    PROC Decorar_Ing165(PERS wobjdata WO_Pastel)
        Mover_en_vacio;
        MoveJ Target_Home_10,Vel_Vacio_Rap,Z_Vacio_Rap,Prototipo_JSDaleman\WObj:=wobj0;
        ReiniciarIndices;
        path_contacto_actual:="p_contacto_165";
        path_vacio_actual:="p_vacio_165";
        Path_Tapa_165ing WO_Pastel;
        Mover_en_vacio;
        MoveJ Target_Home_10,Vel_Vacio_Rap,Z_Vacio_Rap,Prototipo_JSDaleman\WObj:=wobj0;
    ENDPROC
    PROC Path_Tapa_165ing(PERS wobjdata WO_Pastel)
        Path_vacio_ejecucion p_vacio_165, 1, WO_Pastel, FALSE;
        Path_contacto_ejecucion p_contacto_165, 1, 7, WO_Pastel, TRUE;
        Path_vacio_ejecucion p_vacio_165, 2, WO_Pastel, FALSE;
        index_vacio_destino:=15;
        Path_contacto_ejecucion p_contacto_165, 8, 10, WO_Pastel, FALSE;
        Mover_en_contacto;
        TriggC p_contacto_165{11},p_contacto_165{12},Vel_Proceso,triggContactoCir,Z_Proceso,Prototipo_JSDaleman\WObj:=WO_Pastel;
        TriggC p_contacto_165{13},p_contacto_165{14},Vel_Proceso,triggContactoCir,Z_Proceso,Prototipo_JSDaleman\WObj:=WO_Pastel;
        Mover_a_vacio;
        TriggL p_contacto_165{15},Vel_Acercamiento,triggContacto,Z_Acercamiento,Prototipo_JSDaleman\WObj:=WO_Pastel;
        Path_vacio_ejecucion p_vacio_165, 3, WO_Pastel, FALSE;
        index_vacio_destino:=21;
        Mover_a_contacto;
        TriggL p_contacto_165{16},Vel_Acercamiento,triggContacto,Z_Acercamiento,Prototipo_JSDaleman\WObj:=WO_Pastel;
        Mover_en_contacto;
        TriggC p_contacto_165{17},p_contacto_165{18},Vel_Proceso,triggContactoCir,Z_Proceso,Prototipo_JSDaleman\WObj:=WO_Pastel;
        TriggC p_contacto_165{19},p_contacto_165{20},Vel_Proceso,triggContactoCir,Z_Proceso,Prototipo_JSDaleman\WObj:=WO_Pastel;
        Mover_a_vacio;
        TriggL p_contacto_165{21},Vel_Acercamiento,triggContacto,Z_Acercamiento,Prototipo_JSDaleman\WObj:=WO_Pastel;
        Path_vacio_ejecucion p_vacio_165, 4, WO_Pastel, FALSE;
        index_vacio_destino:=28;
        Path_contacto_ejecucion p_contacto_165, 22, 23, WO_Pastel, FALSE;
        Mover_en_contacto;
        TriggC p_contacto_165{24},p_contacto_165{25},Vel_Proceso,triggContactoCir,Z_Proceso,Prototipo_JSDaleman\WObj:=WO_Pastel;
        TriggL p_contacto_165{26},Vel_Proceso,triggContacto,Z_Proceso,Prototipo_JSDaleman\WObj:=WO_Pastel;
        TriggL p_contacto_165{27},Vel_Proceso,triggContacto,Z_Proceso,Prototipo_JSDaleman\WObj:=WO_Pastel;
        Mover_a_vacio;
        TriggL p_contacto_165{28},Vel_Acercamiento,triggContacto,Z_Acercamiento,Prototipo_JSDaleman\WObj:=WO_Pastel;
        Path_vacio_ejecucion p_vacio_165, 5, WO_Pastel, FALSE;
        Path_contacto_ejecucion p_contacto_165, 29, 31, WO_Pastel, TRUE;
        Path_vacio_ejecucion p_vacio_165, 6, WO_Pastel, FALSE;
        Path_contacto_ejecucion p_contacto_165, 32, 39, WO_Pastel, TRUE;
        Path_vacio_ejecucion p_vacio_165, 7, WO_Pastel, FALSE;
        index_vacio_destino:=47;
        Path_contacto_ejecucion p_contacto_165, 40, 42, WO_Pastel, FALSE;
        Mover_en_contacto;
        TriggC p_contacto_165{43},p_contacto_165{44},Vel_Proceso,triggContactoCir,Z_Proceso,Prototipo_JSDaleman\WObj:=WO_Pastel;
        TriggC p_contacto_165{45},p_contacto_165{46},Vel_Proceso,triggContactoCir,Z_Proceso,Prototipo_JSDaleman\WObj:=WO_Pastel;
        Mover_a_vacio;
        TriggL p_contacto_165{47},Vel_Acercamiento,triggContacto,Z_Acercamiento,Prototipo_JSDaleman\WObj:=WO_Pastel;
        Path_vacio_ejecucion p_vacio_165, 8, WO_Pastel, FALSE;
        index_vacio_destino:=55;
        Path_contacto_ejecucion p_contacto_165, 48, 50, WO_Pastel, FALSE;
        Mover_en_contacto;
        TriggC p_contacto_165{51},p_contacto_165{52},Vel_Proceso,triggContactoCir,Z_Proceso,Prototipo_JSDaleman\WObj:=WO_Pastel;
        TriggC p_contacto_165{53},p_contacto_165{54},Vel_Proceso,triggContactoCir,Z_Proceso,Prototipo_JSDaleman\WObj:=WO_Pastel;
        Mover_a_vacio;
        TriggL p_contacto_165{55},Vel_Acercamiento,triggContacto,Z_Acercamiento,Prototipo_JSDaleman\WObj:=WO_Pastel;
        Path_vacio_ejecucion p_vacio_165, 9, WO_Pastel, FALSE;
        index_vacio_destino:=63;
        Path_contacto_ejecucion p_contacto_165, 56, 58, WO_Pastel, FALSE;
        Mover_en_contacto;
        TriggC p_contacto_165{59},p_contacto_165{60},Vel_Proceso,triggContactoCir,Z_Proceso,Prototipo_JSDaleman\WObj:=WO_Pastel;
        TriggC p_contacto_165{61},p_contacto_165{62},Vel_Proceso,triggContactoCir,Z_Proceso,Prototipo_JSDaleman\WObj:=WO_Pastel;
        Mover_a_vacio;
        TriggL p_contacto_165{63},Vel_Acercamiento,triggContacto,Z_Acercamiento,Prototipo_JSDaleman\WObj:=WO_Pastel;
        Path_vacio_ejecucion p_vacio_165, 10, WO_Pastel, FALSE;
        index_vacio_destino:=70;
        Mover_a_contacto;
        TriggL p_contacto_165{64},Vel_Acercamiento,triggContacto,Z_Acercamiento,Prototipo_JSDaleman\WObj:=WO_Pastel;
        Mover_en_contacto;
        TriggC p_contacto_165{65},p_contacto_165{66},Vel_Proceso,triggContactoCir,Z_Proceso,Prototipo_JSDaleman\WObj:=WO_Pastel;
        TriggC p_contacto_165{67},p_contacto_165{68},Vel_Proceso,triggContactoCir,Z_Proceso,Prototipo_JSDaleman\WObj:=WO_Pastel;
        TriggL p_contacto_165{69},Vel_Proceso,triggContacto,Z_Proceso,Prototipo_JSDaleman\WObj:=WO_Pastel;
        Mover_a_vacio;
        TriggL p_contacto_165{70},Vel_Acercamiento,triggContacto,Z_Acercamiento,Prototipo_JSDaleman\WObj:=WO_Pastel;
        Path_vacio_ejecucion p_vacio_165, 11, WO_Pastel, FALSE;
        Path_contacto_ejecucion p_contacto_165, 71, 73, WO_Pastel, TRUE;
        Path_vacio_ejecucion p_vacio_165, 12, WO_Pastel, FALSE;
        index_vacio_destino:=80;
        Path_contacto_ejecucion p_contacto_165, 74, 76, WO_Pastel, FALSE;
        Mover_en_contacto;
        TriggC p_contacto_165{77},p_contacto_165{78},Vel_Proceso,triggContactoCir,Z_Proceso,Prototipo_JSDaleman\WObj:=WO_Pastel;
        TriggL p_contacto_165{79},Vel_Proceso,triggContacto,Z_Proceso,Prototipo_JSDaleman\WObj:=WO_Pastel;
        Mover_a_vacio;
        TriggL p_contacto_165{80},Vel_Acercamiento,triggContacto,Z_Acercamiento,Prototipo_JSDaleman\WObj:=WO_Pastel;
        Path_vacio_ejecucion p_vacio_165, 13, WO_Pastel, FALSE;
        index_vacio_destino:=90;
        Mover_a_contacto;
        TriggL p_contacto_165{81},Vel_Acercamiento,triggContacto,Z_Acercamiento,Prototipo_JSDaleman\WObj:=WO_Pastel;
        Mover_en_contacto;
        TriggC p_contacto_165{82},p_contacto_165{83},Vel_Proceso,triggContactoCir,Z_Proceso,Prototipo_JSDaleman\WObj:=WO_Pastel;
        TriggL p_contacto_165{84},Vel_Proceso,triggContacto,Z_Proceso,Prototipo_JSDaleman\WObj:=WO_Pastel;
        TriggL p_contacto_165{85},Vel_Proceso,triggContacto,Z_Proceso,Prototipo_JSDaleman\WObj:=WO_Pastel;
        TriggC p_contacto_165{86},p_contacto_165{87},Vel_Proceso,triggContactoCir,Z_Proceso,Prototipo_JSDaleman\WObj:=WO_Pastel;
        TriggC p_contacto_165{88},p_contacto_165{89},Vel_Proceso,triggContactoCir,Z_Proceso,Prototipo_JSDaleman\WObj:=WO_Pastel;
        Mover_a_vacio;
        TriggL p_contacto_165{90},Vel_Acercamiento,triggContacto,Z_Acercamiento,Prototipo_JSDaleman\WObj:=WO_Pastel;
        Path_vacio_ejecucion p_vacio_165, 14, WO_Pastel, FALSE;
        index_vacio_destino:=97;
        Mover_a_contacto;
        TriggL p_contacto_165{91},Vel_Acercamiento,triggContacto,Z_Acercamiento,Prototipo_JSDaleman\WObj:=WO_Pastel;
        Mover_en_contacto;
        TriggC p_contacto_165{92},p_contacto_165{93},Vel_Proceso,triggContactoCir,Z_Proceso,Prototipo_JSDaleman\WObj:=WO_Pastel;
        TriggC p_contacto_165{94},p_contacto_165{95},Vel_Proceso,triggContactoCir,Z_Proceso,Prototipo_JSDaleman\WObj:=WO_Pastel;
        TriggL p_contacto_165{96},Vel_Proceso,triggContacto,Z_Proceso,Prototipo_JSDaleman\WObj:=WO_Pastel;
        Mover_a_vacio;
        TriggL p_contacto_165{97},Vel_Acercamiento,triggContacto,Z_Acercamiento,Prototipo_JSDaleman\WObj:=WO_Pastel;
        Path_vacio_ejecucion p_vacio_165, 15, WO_Pastel, FALSE;
        index_vacio_destino:=104;
        Path_contacto_ejecucion p_contacto_165, 98, 100, WO_Pastel, FALSE;
        Mover_en_contacto;
        TriggC p_contacto_165{101},p_contacto_165{102},Vel_Proceso,triggContactoCir,Z_Proceso,Prototipo_JSDaleman\WObj:=WO_Pastel;
        TriggL p_contacto_165{103},Vel_Proceso,triggContacto,Z_Proceso,Prototipo_JSDaleman\WObj:=WO_Pastel;
        Mover_a_vacio;
        TriggL p_contacto_165{104},Vel_Acercamiento,triggContacto,Z_Acercamiento,Prototipo_JSDaleman\WObj:=WO_Pastel;
        Path_vacio_ejecucion p_vacio_165, 16, WO_Pastel, FALSE;
        Path_contacto_ejecucion p_contacto_165, 105, 107, WO_Pastel, TRUE;
        Path_vacio_ejecucion p_vacio_165, 17, WO_Pastel, FALSE;
        Path_contacto_ejecucion p_contacto_165, 108, 109, WO_Pastel, TRUE;
        Path_vacio_ejecucion p_vacio_165, 18, WO_Pastel, FALSE;
        index_vacio_destino:=116;
        Mover_a_contacto;
        TriggL p_contacto_165{110},Vel_Acercamiento,triggContacto,Z_Acercamiento,Prototipo_JSDaleman\WObj:=WO_Pastel;
        Mover_en_contacto;
        TriggC p_contacto_165{111},p_contacto_165{112},Vel_Proceso,triggContactoCir,Z_Proceso,Prototipo_JSDaleman\WObj:=WO_Pastel;
        TriggC p_contacto_165{113},p_contacto_165{114},Vel_Proceso,triggContactoCir,Z_Proceso,Prototipo_JSDaleman\WObj:=WO_Pastel;
        TriggL p_contacto_165{115},Vel_Proceso,triggContacto,Z_Proceso,Prototipo_JSDaleman\WObj:=WO_Pastel;
        Mover_a_vacio;
        TriggL p_contacto_165{116},Vel_Acercamiento,triggContacto,Z_Acercamiento,Prototipo_JSDaleman\WObj:=WO_Pastel;
        Path_vacio_ejecucion p_vacio_165, 19, WO_Pastel, FALSE;
        Path_contacto_ejecucion p_contacto_165, 117, 121, WO_Pastel, TRUE;
        Path_vacio_ejecucion p_vacio_165, 20, WO_Pastel, FALSE;
        Path_contacto_ejecucion p_contacto_165, 122, 124, WO_Pastel, TRUE;
        Path_vacio_ejecucion p_vacio_165, 21, WO_Pastel, FALSE;
        Path_contacto_ejecucion p_contacto_165, 125, 127, WO_Pastel, TRUE;
        Path_vacio_ejecucion p_vacio_165, 22, WO_Pastel, FALSE;
        index_vacio_destino:=135;
        Path_contacto_ejecucion p_contacto_165, 128, 130, WO_Pastel, FALSE;
        Mover_en_contacto;
        TriggC p_contacto_165{131},p_contacto_165{132},Vel_Proceso,triggContactoCir,Z_Proceso,Prototipo_JSDaleman\WObj:=WO_Pastel;
        TriggC p_contacto_165{133},p_contacto_165{134},Vel_Proceso,triggContactoCir,Z_Proceso,Prototipo_JSDaleman\WObj:=WO_Pastel;
        Mover_a_vacio;
        TriggL p_contacto_165{135},Vel_Acercamiento,triggContacto,Z_Acercamiento,Prototipo_JSDaleman\WObj:=WO_Pastel;
        Path_vacio_ejecucion p_vacio_165, 23, WO_Pastel, FALSE;
        index_vacio_destino:=139;
        Mover_a_contacto;
        TriggL p_contacto_165{136},Vel_Acercamiento,triggContacto,Z_Acercamiento,Prototipo_JSDaleman\WObj:=WO_Pastel;
        Mover_en_contacto;
        TriggC p_contacto_165{137},p_contacto_165{138},Vel_Proceso,triggContactoCir,Z_Proceso,Prototipo_JSDaleman\WObj:=WO_Pastel;
        Mover_a_vacio;
        TriggL p_contacto_165{139},Vel_Acercamiento,triggContacto,Z_Acercamiento,Prototipo_JSDaleman\WObj:=WO_Pastel;
        Path_vacio_ejecucion p_vacio_165, 24, WO_Pastel, FALSE;
        index_vacio_destino:=143;
        Mover_a_contacto;
        TriggL p_contacto_165{140},Vel_Acercamiento,triggContacto,Z_Acercamiento,Prototipo_JSDaleman\WObj:=WO_Pastel;
        Mover_en_contacto;
        TriggC p_contacto_165{141},p_contacto_165{142},Vel_Proceso,triggContactoCir,Z_Proceso,Prototipo_JSDaleman\WObj:=WO_Pastel;
        Mover_a_vacio;
        TriggL p_contacto_165{143},Vel_Acercamiento,triggContacto,Z_Acercamiento,Prototipo_JSDaleman\WObj:=WO_Pastel;
        Path_vacio_ejecucion p_vacio_165, 25, WO_Pastel, FALSE;
        index_vacio_destino:=147;
        Mover_a_contacto;
        TriggL p_contacto_165{144},Vel_Acercamiento,triggContacto,Z_Acercamiento,Prototipo_JSDaleman\WObj:=WO_Pastel;
        Mover_en_contacto;
        TriggC p_contacto_165{145},p_contacto_165{146},Vel_Proceso,triggContactoCir,Z_Proceso,Prototipo_JSDaleman\WObj:=WO_Pastel;
        Mover_a_vacio;
        TriggL p_contacto_165{147},Vel_Acercamiento,triggContacto,Z_Acercamiento,Prototipo_JSDaleman\WObj:=WO_Pastel;
        Path_vacio_ejecucion p_vacio_165, 26, WO_Pastel, FALSE;
        Path_contacto_ejecucion p_contacto_165, 148, 150, WO_Pastel, TRUE;
        Path_vacio_ejecucion p_vacio_165, 27, WO_Pastel, FALSE;
        index_vacio_destino:=154;
        Mover_a_contacto;
        TriggL p_contacto_165{151},Vel_Acercamiento,triggContacto,Z_Acercamiento,Prototipo_JSDaleman\WObj:=WO_Pastel;
        Mover_en_contacto;
        TriggC p_contacto_165{152},p_contacto_165{153},Vel_Proceso,triggContactoCir,Z_Proceso,Prototipo_JSDaleman\WObj:=WO_Pastel;
        Mover_a_vacio;
        TriggL p_contacto_165{154},Vel_Acercamiento,triggContacto,Z_Acercamiento,Prototipo_JSDaleman\WObj:=WO_Pastel;
        Path_vacio_ejecucion p_vacio_165, 28, WO_Pastel, FALSE;
        index_vacio_destino:=158;
        Mover_a_contacto;
        TriggL p_contacto_165{155},Vel_Acercamiento,triggContacto,Z_Acercamiento,Prototipo_JSDaleman\WObj:=WO_Pastel;
        Mover_en_contacto;
        TriggC p_contacto_165{156},p_contacto_165{157},Vel_Proceso,triggContactoCir,Z_Proceso,Prototipo_JSDaleman\WObj:=WO_Pastel;
        Mover_a_vacio;
        TriggL p_contacto_165{158},Vel_Acercamiento,triggContacto,Z_Acercamiento,Prototipo_JSDaleman\WObj:=WO_Pastel;
        Path_vacio_ejecucion p_vacio_165, 29, WO_Pastel, FALSE;
        index_vacio_destino:=162;
        Mover_a_contacto;
        TriggL p_contacto_165{159},Vel_Acercamiento,triggContacto,Z_Acercamiento,Prototipo_JSDaleman\WObj:=WO_Pastel;
        Mover_en_contacto;
        TriggC p_contacto_165{160},p_contacto_165{161},Vel_Proceso,triggContactoCir,Z_Proceso,Prototipo_JSDaleman\WObj:=WO_Pastel;
        Mover_a_vacio;
        TriggL p_contacto_165{162},Vel_Acercamiento,triggContacto,Z_Acercamiento,Prototipo_JSDaleman\WObj:=WO_Pastel;
        Path_vacio_ejecucion p_vacio_165, 30, WO_Pastel, FALSE;
        index_vacio_destino:=170;
        Path_contacto_ejecucion p_contacto_165, 163, 165, WO_Pastel, FALSE;
        Mover_en_contacto;
        TriggC p_contacto_165{166},p_contacto_165{167},Vel_Proceso,triggContactoCir,Z_Proceso,Prototipo_JSDaleman\WObj:=WO_Pastel;
        TriggC p_contacto_165{168},p_contacto_165{169},Vel_Proceso,triggContactoCir,Z_Proceso,Prototipo_JSDaleman\WObj:=WO_Pastel;
        Mover_a_vacio;
        TriggL p_contacto_165{170},Vel_Acercamiento,triggContacto,Z_Acercamiento,Prototipo_JSDaleman\WObj:=WO_Pastel;
        Path_vacio_ejecucion p_vacio_165, 31, WO_Pastel, FALSE;
        index_vacio_destino:=178;
        Path_contacto_ejecucion p_contacto_165, 171, 173, WO_Pastel, FALSE;
        Mover_en_contacto;
        TriggC p_contacto_165{174},p_contacto_165{175},Vel_Proceso,triggContactoCir,Z_Proceso,Prototipo_JSDaleman\WObj:=WO_Pastel;
        TriggL p_contacto_165{176},Vel_Proceso,triggContacto,Z_Proceso,Prototipo_JSDaleman\WObj:=WO_Pastel;
        TriggL p_contacto_165{177},Vel_Proceso,triggContacto,Z_Proceso,Prototipo_JSDaleman\WObj:=WO_Pastel;
        Mover_a_vacio;
        TriggL p_contacto_165{178},Vel_Acercamiento,triggContacto,Z_Acercamiento,Prototipo_JSDaleman\WObj:=WO_Pastel;
        Path_vacio_ejecucion p_vacio_165, 32, WO_Pastel, FALSE;
        index_vacio_destino:=184;
        Mover_a_contacto;
        TriggL p_contacto_165{179},Vel_Acercamiento,triggContacto,Z_Acercamiento,Prototipo_JSDaleman\WObj:=WO_Pastel;
        Mover_en_contacto;
        TriggC p_contacto_165{180},p_contacto_165{181},Vel_Proceso,triggContactoCir,Z_Proceso,Prototipo_JSDaleman\WObj:=WO_Pastel;
        TriggC p_contacto_165{182},p_contacto_165{183},Vel_Proceso,triggContactoCir,Z_Proceso,Prototipo_JSDaleman\WObj:=WO_Pastel;
        Mover_a_vacio;
        TriggL p_contacto_165{184},Vel_Acercamiento,triggContacto,Z_Acercamiento,Prototipo_JSDaleman\WObj:=WO_Pastel;
        Path_vacio_ejecucion p_vacio_165, 33, WO_Pastel, FALSE;
        index_vacio_destino:=190;
        Mover_a_contacto;
        TriggL p_contacto_165{185},Vel_Acercamiento,triggContacto,Z_Acercamiento,Prototipo_JSDaleman\WObj:=WO_Pastel;
        Mover_en_contacto;
        TriggC p_contacto_165{186},p_contacto_165{187},Vel_Proceso,triggContactoCir,Z_Proceso,Prototipo_JSDaleman\WObj:=WO_Pastel;
        TriggC p_contacto_165{188},p_contacto_165{189},Vel_Proceso,triggContactoCir,Z_Proceso,Prototipo_JSDaleman\WObj:=WO_Pastel;
        Mover_a_vacio;
        TriggL p_contacto_165{190},Vel_Acercamiento,triggContacto,Z_Acercamiento,Prototipo_JSDaleman\WObj:=WO_Pastel;
        Path_vacio_ejecucion p_vacio_165, 34, WO_Pastel, FALSE;
        index_vacio_destino:=198;
        Mover_a_contacto;
        TriggL p_contacto_165{191},Vel_Acercamiento,triggContacto,Z_Acercamiento,Prototipo_JSDaleman\WObj:=WO_Pastel;
        Mover_en_contacto;
        TriggC p_contacto_165{192},p_contacto_165{193},Vel_Proceso,triggContactoCir,Z_Proceso,Prototipo_JSDaleman\WObj:=WO_Pastel;
        TriggL p_contacto_165{194},Vel_Proceso,triggContacto,Z_Proceso,Prototipo_JSDaleman\WObj:=WO_Pastel;
        TriggL p_contacto_165{195},Vel_Proceso,triggContacto,Z_Proceso,Prototipo_JSDaleman\WObj:=WO_Pastel;
        TriggC p_contacto_165{196},p_contacto_165{197},Vel_Proceso,triggContactoCir,Z_Proceso,Prototipo_JSDaleman\WObj:=WO_Pastel;
        Mover_a_vacio;
        TriggL p_contacto_165{198},Vel_Acercamiento,triggContacto,Z_Acercamiento,Prototipo_JSDaleman\WObj:=WO_Pastel;
        Path_vacio_ejecucion p_vacio_165, 35, WO_Pastel, FALSE;
        Path_contacto_ejecucion p_contacto_165, 199, 201, WO_Pastel, TRUE;
        Path_vacio_ejecucion p_vacio_165, 36, WO_Pastel, FALSE;
        Path_contacto_ejecucion p_contacto_165, 202, 204, WO_Pastel, TRUE;
        Path_vacio_ejecucion p_vacio_165, 37, WO_Pastel, FALSE;
        Path_contacto_ejecucion p_contacto_165, 205, 207, WO_Pastel, TRUE;
        Path_vacio_ejecucion p_vacio_165, 38, WO_Pastel, FALSE;
        Path_contacto_ejecucion p_contacto_165, 208, 210, WO_Pastel, TRUE;
        Path_vacio_ejecucion p_vacio_165, 39, WO_Pastel, FALSE;
        index_vacio_destino:=214;
        Mover_a_contacto;
        TriggL p_contacto_165{211},Vel_Acercamiento,triggContacto,Z_Acercamiento,Prototipo_JSDaleman\WObj:=WO_Pastel;
        Mover_en_contacto;
        TriggC p_contacto_165{212},p_contacto_165{213},Vel_Proceso,triggContactoCir,Z_Proceso,Prototipo_JSDaleman\WObj:=WO_Pastel;
        Mover_a_vacio;
        TriggL p_contacto_165{214},Vel_Acercamiento,triggContacto,Z_Acercamiento,Prototipo_JSDaleman\WObj:=WO_Pastel;
        Path_vacio_ejecucion p_vacio_165, 40, WO_Pastel, FALSE;
        index_vacio_destino:=218;
        Mover_a_contacto;
        TriggL p_contacto_165{215},Vel_Acercamiento,triggContacto,Z_Acercamiento,Prototipo_JSDaleman\WObj:=WO_Pastel;
        Mover_en_contacto;
        TriggC p_contacto_165{216},p_contacto_165{217},Vel_Proceso,triggContactoCir,Z_Proceso,Prototipo_JSDaleman\WObj:=WO_Pastel;
        Mover_a_vacio;
        TriggL p_contacto_165{218},Vel_Acercamiento,triggContacto,Z_Acercamiento,Prototipo_JSDaleman\WObj:=WO_Pastel;
        Path_vacio_ejecucion p_vacio_165, 41, WO_Pastel, FALSE;
        index_vacio_destino:=222;
        Mover_a_contacto;
        TriggL p_contacto_165{219},Vel_Acercamiento,triggContacto,Z_Acercamiento,Prototipo_JSDaleman\WObj:=WO_Pastel;
        Mover_en_contacto;
        TriggC p_contacto_165{220},p_contacto_165{221},Vel_Proceso,triggContactoCir,Z_Proceso,Prototipo_JSDaleman\WObj:=WO_Pastel;
        Mover_a_vacio;
        TriggL p_contacto_165{222},Vel_Acercamiento,triggContacto,Z_Acercamiento,Prototipo_JSDaleman\WObj:=WO_Pastel;
        Path_vacio_ejecucion p_vacio_165, 42, WO_Pastel, FALSE;
        index_vacio_destino:=227;
        Mover_a_contacto;
        TriggL p_contacto_165{223},Vel_Acercamiento,triggContacto,Z_Acercamiento,Prototipo_JSDaleman\WObj:=WO_Pastel;
        Mover_en_contacto;
        TriggC p_contacto_165{224},p_contacto_165{225},Vel_Proceso,triggContactoCir,Z_Proceso,Prototipo_JSDaleman\WObj:=WO_Pastel;
        TriggL p_contacto_165{226},Vel_Proceso,triggContacto,Z_Proceso,Prototipo_JSDaleman\WObj:=WO_Pastel;
        Mover_a_vacio;
        TriggL p_contacto_165{227},Vel_Acercamiento,triggContacto,Z_Acercamiento,Prototipo_JSDaleman\WObj:=WO_Pastel;
        Path_vacio_ejecucion p_vacio_165, 43, WO_Pastel, FALSE;
        index_vacio_destino:=232;
        Mover_a_contacto;
        TriggL p_contacto_165{228},Vel_Acercamiento,triggContacto,Z_Acercamiento,Prototipo_JSDaleman\WObj:=WO_Pastel;
        TriggL p_contacto_165{229},Vel_Proceso,triggContacto,Z_Proceso,Prototipo_JSDaleman\WObj:=WO_Pastel;
        TriggC p_contacto_165{230},p_contacto_165{231},Vel_Proceso,triggContactoCir,Z_Proceso,Prototipo_JSDaleman\WObj:=WO_Pastel;
        Mover_a_vacio;
        TriggL p_contacto_165{232},Vel_Acercamiento,triggContacto,Z_Acercamiento,Prototipo_JSDaleman\WObj:=WO_Pastel;
        Path_vacio_ejecucion p_vacio_165, 44, WO_Pastel, FALSE;
        index_vacio_destino:=236;
        Mover_a_contacto;
        TriggL p_contacto_165{233},Vel_Acercamiento,triggContacto,Z_Acercamiento,Prototipo_JSDaleman\WObj:=WO_Pastel;
        Mover_en_contacto;
        TriggC p_contacto_165{234},p_contacto_165{235},Vel_Proceso,triggContactoCir,Z_Proceso,Prototipo_JSDaleman\WObj:=WO_Pastel;
        Mover_a_vacio;
        TriggL p_contacto_165{236},Vel_Acercamiento,triggContacto,Z_Acercamiento,Prototipo_JSDaleman\WObj:=WO_Pastel;
        Path_vacio_ejecucion p_vacio_165, 45, WO_Pastel, FALSE;
        index_vacio_destino:=240;
        Mover_a_contacto;
        TriggL p_contacto_165{237},Vel_Acercamiento,triggContacto,Z_Acercamiento,Prototipo_JSDaleman\WObj:=WO_Pastel;
        Mover_en_contacto;
        TriggC p_contacto_165{238},p_contacto_165{239},Vel_Proceso,triggContactoCir,Z_Proceso,Prototipo_JSDaleman\WObj:=WO_Pastel;
        Mover_a_vacio;
        TriggL p_contacto_165{240},Vel_Acercamiento,triggContacto,Z_Acercamiento,Prototipo_JSDaleman\WObj:=WO_Pastel;
        Path_vacio_ejecucion p_vacio_165, 46, WO_Pastel, FALSE;
        index_vacio_destino:=244;
        Mover_a_contacto;
        TriggL p_contacto_165{241},Vel_Acercamiento,triggContacto,Z_Acercamiento,Prototipo_JSDaleman\WObj:=WO_Pastel;
        Mover_en_contacto;
        TriggC p_contacto_165{242},p_contacto_165{243},Vel_Proceso,triggContactoCir,Z_Proceso,Prototipo_JSDaleman\WObj:=WO_Pastel;
        Mover_a_vacio;
        TriggL p_contacto_165{244},Vel_Acercamiento,triggContacto,Z_Acercamiento,Prototipo_JSDaleman\WObj:=WO_Pastel;
        Path_vacio_ejecucion p_vacio_165, 47, WO_Pastel, FALSE;
        index_vacio_destino:=247;
        Mover_a_contacto;
        TriggL p_contacto_165{245},Vel_Acercamiento,triggContacto,Z_Acercamiento,Prototipo_JSDaleman\WObj:=WO_Pastel;
        Mover_en_contacto;
        TriggL p_contacto_165{246},Vel_Proceso,triggContacto,Z_Proceso,Prototipo_JSDaleman\WObj:=WO_Pastel;
        Mover_a_vacio;
        TriggL p_contacto_165{247},Vel_Acercamiento,triggContacto,Z_Acercamiento,Prototipo_JSDaleman\WObj:=WO_Pastel;
        Path_vacio_ejecucion p_vacio_165, 48, WO_Pastel, FALSE;
        Path_contacto_ejecucion p_contacto_165, 248, 250, WO_Pastel, TRUE;
        Path_vacio_ejecucion p_vacio_165, 49, WO_Pastel, FALSE;
        Path_contacto_ejecucion p_contacto_165, 251, 253, WO_Pastel, TRUE;
        Path_vacio_ejecucion p_vacio_165, 50, WO_Pastel, FALSE;
        Path_contacto_ejecucion p_contacto_165, 254, 256, WO_Pastel, TRUE;
        Path_vacio_ejecucion p_vacio_165, 51, WO_Pastel, FALSE;
        Path_contacto_ejecucion p_contacto_165, 257, 259, WO_Pastel, TRUE;
        Path_vacio_ejecucion p_vacio_165, 52, WO_Pastel, FALSE;
        Path_contacto_ejecucion p_contacto_165, 260, 262, WO_Pastel, TRUE;
        Path_vacio_ejecucion p_vacio_165, 53, WO_Pastel, FALSE;
        Path_contacto_ejecucion p_contacto_165, 263, 266, WO_Pastel, TRUE;
        Path_vacio_ejecucion p_vacio_165, 54, WO_Pastel, FALSE;
        index_vacio_destino:=276;
        Mover_a_contacto;
        TriggL p_contacto_165{267},Vel_Acercamiento,triggContacto,Z_Acercamiento,Prototipo_JSDaleman\WObj:=WO_Pastel;
        Mover_en_contacto;
        TriggC p_contacto_165{268},p_contacto_165{269},Vel_Proceso,triggContactoCir,Z_Proceso,Prototipo_JSDaleman\WObj:=WO_Pastel;
        TriggC p_contacto_165{270},p_contacto_165{271},Vel_Proceso,triggContactoCir,Z_Proceso,Prototipo_JSDaleman\WObj:=WO_Pastel;
        TriggC p_contacto_165{272},p_contacto_165{273},Vel_Proceso,triggContactoCir,Z_Proceso,Prototipo_JSDaleman\WObj:=WO_Pastel;
        TriggC p_contacto_165{274},p_contacto_165{275},Vel_Proceso,triggContactoCir,Z_Proceso,Prototipo_JSDaleman\WObj:=WO_Pastel;
        Mover_a_vacio;
        TriggL p_contacto_165{276},Vel_Acercamiento,triggContacto,Z_Acercamiento,Prototipo_JSDaleman\WObj:=WO_Pastel;
        Path_vacio_ejecucion p_vacio_165, 55, WO_Pastel, FALSE;
        index_vacio_destino:=285;
        Mover_a_contacto;
        TriggL p_contacto_165{277},Vel_Acercamiento,triggContacto,Z_Acercamiento,Prototipo_JSDaleman\WObj:=WO_Pastel;
        Mover_en_contacto;
        TriggC p_contacto_165{278},p_contacto_165{279},Vel_Proceso,triggContactoCir,Z_Proceso,Prototipo_JSDaleman\WObj:=WO_Pastel;
        TriggL p_contacto_165{280},Vel_Proceso,triggContacto,Z_Proceso,Prototipo_JSDaleman\WObj:=WO_Pastel;
        TriggC p_contacto_165{281},p_contacto_165{282},Vel_Proceso,triggContactoCir,Z_Proceso,Prototipo_JSDaleman\WObj:=WO_Pastel;
        TriggC p_contacto_165{283},p_contacto_165{284},Vel_Proceso,triggContactoCir,Z_Proceso,Prototipo_JSDaleman\WObj:=WO_Pastel;
        Mover_a_vacio;
        TriggL p_contacto_165{285},Vel_Acercamiento,triggContacto,Z_Acercamiento,Prototipo_JSDaleman\WObj:=WO_Pastel;
        Path_vacio_ejecucion p_vacio_165, 56, WO_Pastel, FALSE;
        Path_contacto_ejecucion p_contacto_165, 286, 289, WO_Pastel, TRUE;
        Path_vacio_ejecucion p_vacio_165, 57, WO_Pastel, FALSE;
        Path_contacto_ejecucion p_contacto_165, 290, 292, WO_Pastel, TRUE;
        Path_vacio_ejecucion p_vacio_165, 58, WO_Pastel, FALSE;
        index_vacio_destino:=298;
        Mover_a_contacto;
        TriggL p_contacto_165{293},Vel_Acercamiento,triggContacto,Z_Acercamiento,Prototipo_JSDaleman\WObj:=WO_Pastel;
        Mover_en_contacto;
        TriggC p_contacto_165{294},p_contacto_165{295},Vel_Proceso,triggContactoCir,Z_Proceso,Prototipo_JSDaleman\WObj:=WO_Pastel;
        TriggL p_contacto_165{296},Vel_Proceso,triggContacto,Z_Proceso,Prototipo_JSDaleman\WObj:=WO_Pastel;
        TriggL p_contacto_165{297},Vel_Proceso,triggContacto,Z_Proceso,Prototipo_JSDaleman\WObj:=WO_Pastel;
        Mover_a_vacio;
        TriggL p_contacto_165{298},Vel_Acercamiento,triggContacto,Z_Acercamiento,Prototipo_JSDaleman\WObj:=WO_Pastel;
        Path_vacio_ejecucion p_vacio_165, 59, WO_Pastel, FALSE;
        index_vacio_destino:=304;
        Mover_a_contacto;
        TriggL p_contacto_165{299},Vel_Acercamiento,triggContacto,Z_Acercamiento,Prototipo_JSDaleman\WObj:=WO_Pastel;
        Mover_en_contacto;
        TriggC p_contacto_165{300},p_contacto_165{301},Vel_Proceso,triggContactoCir,Z_Proceso,Prototipo_JSDaleman\WObj:=WO_Pastel;
        TriggC p_contacto_165{302},p_contacto_165{303},Vel_Proceso,triggContactoCir,Z_Proceso,Prototipo_JSDaleman\WObj:=WO_Pastel;
        Mover_a_vacio;
        TriggL p_contacto_165{304},Vel_Acercamiento,triggContacto,Z_Acercamiento,Prototipo_JSDaleman\WObj:=WO_Pastel;
        Path_vacio_ejecucion p_vacio_165, 60, WO_Pastel, FALSE;
        index_vacio_destino:=310;
        Mover_a_contacto;
        TriggL p_contacto_165{305},Vel_Acercamiento,triggContacto,Z_Acercamiento,Prototipo_JSDaleman\WObj:=WO_Pastel;
        Mover_en_contacto;
        TriggC p_contacto_165{306},p_contacto_165{307},Vel_Proceso,triggContactoCir,Z_Proceso,Prototipo_JSDaleman\WObj:=WO_Pastel;
        TriggL p_contacto_165{308},Vel_Proceso,triggContacto,Z_Proceso,Prototipo_JSDaleman\WObj:=WO_Pastel;
        TriggL p_contacto_165{309},Vel_Proceso,triggContacto,Z_Proceso,Prototipo_JSDaleman\WObj:=WO_Pastel;
        Mover_a_vacio;
        TriggL p_contacto_165{310},Vel_Acercamiento,triggContacto,Z_Acercamiento,Prototipo_JSDaleman\WObj:=WO_Pastel;
        Path_vacio_ejecucion p_vacio_165, 61, WO_Pastel, FALSE;
        index_vacio_destino:=319;
        Mover_a_contacto;
        TriggL p_contacto_165{311},Vel_Acercamiento,triggContacto,Z_Acercamiento,Prototipo_JSDaleman\WObj:=WO_Pastel;
        Mover_en_contacto;
        TriggC p_contacto_165{312},p_contacto_165{313},Vel_Proceso,triggContactoCir,Z_Proceso,Prototipo_JSDaleman\WObj:=WO_Pastel;
        TriggL p_contacto_165{314},Vel_Proceso,triggContacto,Z_Proceso,Prototipo_JSDaleman\WObj:=WO_Pastel;
        TriggC p_contacto_165{315},p_contacto_165{316},Vel_Proceso,triggContactoCir,Z_Proceso,Prototipo_JSDaleman\WObj:=WO_Pastel;
        TriggC p_contacto_165{317},p_contacto_165{318},Vel_Proceso,triggContactoCir,Z_Proceso,Prototipo_JSDaleman\WObj:=WO_Pastel;
        Mover_a_vacio;
        TriggL p_contacto_165{319},Vel_Acercamiento,triggContacto,Z_Acercamiento,Prototipo_JSDaleman\WObj:=WO_Pastel;
    ENDPROC

ENDMODULE

--- Controller Data/IRB140_LabSIR/RAPID/TASK1/PROGMOD/Interrupciones.mod ---
MODULE Interrupciones

    !***********************************************************
    !
    ! Modulo:  Interrupciones
    !
    ! Descripción:
    !   Modulo de manejo de interrupciones para manejo de la HMI
    !
    ! Autor: Juan_Daleman
    !
    ! Versión: 1.0
    !
    !***********************************************************

     !Variables de interrupcion
     VAR intnum DIHomeActiva;
     VAR intnum DIManteActiva;
     VAR intnum DIEsperaActiva;
     VAR intnum BoolHomeActiva;
     VAR intnum BoolTransActiva;
     VAR intnum BoolManteActiva;
     VAR intnum BoolEsperaActiva;
     VAR intnum BoolRevisionActiva;
     VAR intnum ParadaEmergencia;
     VAR intnum PausaContinuar;
     VAR intnum ReiniciarRut;
     VAR intnum IncrementoIndicesContacto;
     VAR intnum IncrementoIndicesContactoCirculo;
     VAR intnum IncrementoIndicesVacio;

     !Variables de mensajes de error para el usuario
     VAR btnres respuesta_parada;
     CONST string mensaje_parada{3} := ["Parada del sistema ejecutada", "Es necesario realizar rearme de operación", "Reinicie el sistema"];

     VAR btnres respuesta_reinicio;
     CONST string mensaje_reinicio{3} := ["Reinicio del sistema ejecutado", "Se reiniciara todo el sistema", "es necesario reiniciar el sistema de supervisión"];

    TRAP Path_Home_DI
        IDelete socket_com_in;
        IDisable;
        StopMove;
        ClearPath;
        StorePath;
        SetDO DO_02,0;
        SetDO DO_03,0;
        Test_Transi:=FALSE;
        StartMove;
        MoveJ Target_Home_10,Vel_Vacio_Rap,Z_Vacio_Rap,Prototipo_JSDaleman\WObj:=wobj0;
        MoveJ Target_Home_20,Vel_Vacio_Rap,Z_Paro,Prototipo_JSDaleman\WObj:=wobj0;
        RestoPath;
        StopMove;
        SetDO DO_01,1;
        IEnable;
        CONNECT socket_com_in WITH SockDataIn;
        IPers cmd, socket_com_in;
    ENDTRAP
    TRAP Path_Home
        IDelete socket_com_in;
        IDisable;
        StopMove;
        ClearPath;
        StorePath;
        SetDO DO_02,0;
        SetDO DO_03,0;
        Test_Transi:=FALSE;
        StartMove;
        IF Bool_Home = TRUE THEN
            MoveJ Target_Home_10,Vel_Vacio_Rap,Z_Vacio_Rap,Prototipo_JSDaleman\WObj:=wobj0;
            MoveJ Target_Home_20,Vel_Vacio_Rap,Z_Paro,Prototipo_JSDaleman\WObj:=wobj0;
            SetDO DO_01,1;
        ENDIF
        RestoPath;
        StopMove;
        IEnable;
        CONNECT socket_com_in WITH SockDataIn;
        IPers cmd, socket_com_in;
    ENDTRAP
    TRAP Path_Transicion_Home
        IDelete socket_com_in;
        IDisable;
        StopMove;
        ClearPath;
        StorePath;
        SetDO DO_01,0;
        SetDO DO_02,0;
        SetDO DO_03,0;
        StartMove;
        IF Bool_Transic = TRUE THEN
            MoveJ Target_Home_10,Vel_Vacio_Rap,Z_Paro,Prototipo_JSDaleman\WObj:=wobj0;
            Test_Transi:=TRUE;
        ENDIF
        RestoPath;
        StopMove;
        IEnable;
        CONNECT socket_com_in WITH SockDataIn;
        IPers cmd, socket_com_in;
    ENDTRAP
    TRAP Path_Mantenimiento_DI
        IDelete socket_com_in;
        IDisable;
        StopMove;
        ClearPath;
        StorePath;
        SetDO DO_01,0;
        SetDO DO_03,0;
        Test_Transi:=FALSE;
        StartMove;
        MoveJ Target_Home_10,Vel_Vacio_Rap,Z_Vacio_Rap,Prototipo_JSDaleman\WObj:=wobj0;
        MoveJ Target_Mantenimiento,Vel_Vacio_Rap,Z_Paro,Prototipo_JSDaleman\WObj:=wobj0;
        SetDO DO_02,1;
        RestoPath;
        StopMove;
        IEnable;
        CONNECT socket_com_in WITH SockDataIn;
        IPers cmd, socket_com_in;
    ENDTRAP
    TRAP Path_Mantenimiento
        IDelete socket_com_in;
        IDisable;
        StopMove;
        ClearPath;
        StorePath;
        SetDO DO_01,0;
        SetDO DO_03,0;
        Test_Transi:=FALSE;
        StartMove;
        IF Bool_Mant = TRUE THEN
            MoveJ Target_Home_10,Vel_Vacio_Rap,Z_Vacio_Rap,Prototipo_JSDaleman\WObj:=wobj0;
            MoveJ Target_Mantenimiento,Vel_Vacio_Rap,Z_Paro,Prototipo_JSDaleman\WObj:=wobj0;
            SetDO DO_02,1;
        ENDIF
        RestoPath;
        StopMove;
        IEnable;
        CONNECT socket_com_in WITH SockDataIn;
        IPers cmd, socket_com_in;
    ENDTRAP
    TRAP Path_IntEspera_DI
        IDelete socket_com_in;
        IDisable;
        StopMove;
        ClearPath;
        StorePath;
        SetDO DO_01,0;
        SetDO DO_02,0;
        SetDO DO_03,0;
        Test_Transi:=FALSE;
        StartMove;
        MoveJ Target_Home_10,Vel_Vacio_Rap,Z_Vacio_Rap,Prototipo_JSDaleman\WObj:=wobj0;
        MoveJ Target_Espera,Vel_Vacio_Rap,Z_Paro,Prototipo_JSDaleman\WObj:=wobj0;
        SetDO DO_03,1;
        RestoPath;
        StopMove;
        IEnable;
        CONNECT socket_com_in WITH SockDataIn;
        IPers cmd, socket_com_in;
    ENDTRAP
    TRAP Path_IntEspera
        IDelete socket_com_in;
        IDisable;
        StopMove;
        ClearPath;
        StorePath;
        SetDO DO_01,0;
        SetDO DO_02,0;
        SetDO DO_03,0;
        Test_Transi:=FALSE;
        StartMove;
        IF Bool_Esper = TRUE THEN
            MoveJ Target_Home_10,Vel_Vacio_Rap,Z_Vacio_Rap,Prototipo_JSDaleman\WObj:=wobj0;
            MoveJ Target_Espera,Vel_Vacio_Rap,Z_Paro,Prototipo_JSDaleman\WObj:=wobj0;
        ENDIF
        SetDO DO_03,1;
        RestoPath;
        StopMove;
        IEnable;
        CONNECT socket_com_in WITH SockDataIn;
        IPers cmd, socket_com_in;
    ENDTRAP
    TRAP Path_PuntosContacto_LabSir
        IDelete socket_com_in;
        IDisable;
        StopMove;
        ClearPath;
        StorePath;
        Test_Transi:=FALSE;
        StartMove;
        IF Bool_RevWO = TRUE THEN
            MoveJ Target_Home_10,Vel_Vacio_Rap,Z_Vacio_Rap,Prototipo_JSDaleman\WObj:=wobj0;
            MoveJ Target_APuntosRef_10,Vel_Vacio_Rap,Z_VacioMov,Prototipo_JSDaleman\WObj:=WO_PastelDef;
            WaitUntil Bool_Confirm=TRUE;
            WaitUntil Bool_Confirm=FALSE;
            MoveL Target_APuntosRef_20,Vel_Acercamiento,Z_Acercamiento,Prototipo_JSDaleman\WObj:=WO_PastelDef;
            WaitUntil Bool_Confirm=TRUE;
            WaitUntil Bool_Confirm=FALSE;
            MoveL Target_APuntosRef_30,Vel_Acercamiento,Z_Acercamiento,Prototipo_JSDaleman\WObj:=WO_PastelDef;
            MoveJ Target_APuntosRef_40,Vel_Vacio,Z_VacioMov,Prototipo_JSDaleman\WObj:=WO_PastelDef;
            WaitUntil Bool_Confirm=TRUE;
            WaitUntil Bool_Confirm=FALSE;
            MoveL Target_APuntosRef_50,Vel_Acercamiento,Z_Acercamiento,Prototipo_JSDaleman\WObj:=WO_PastelDef;
            WaitUntil Bool_Confirm=TRUE;
            WaitUntil Bool_Confirm=FALSE;
            MoveL Target_APuntosRef_60,Vel_Acercamiento,Z_Acercamiento,Prototipo_JSDaleman\WObj:=WO_PastelDef;
            MoveJ Target_APuntosRef_70,Vel_Vacio,Z_VacioMov,Prototipo_JSDaleman\WObj:=WO_PastelDef;
            WaitUntil Bool_Confirm=TRUE;
            WaitUntil Bool_Confirm=FALSE;
            MoveL Target_APuntosRef_80,Vel_Acercamiento,Z_Acercamiento,Prototipo_JSDaleman\WObj:=WO_PastelDef;
            WaitUntil Bool_Confirm=TRUE;
            WaitUntil Bool_Confirm=FALSE;
            MoveL Target_APuntosRef_90,Vel_Acercamiento,Z_Acercamiento,Prototipo_JSDaleman\WObj:=WO_PastelDef;
            MoveJ Target_APuntosRef_100,Vel_Vacio,Z_VacioMov,Prototipo_JSDaleman\WObj:=WO_PastelDef;
            WaitUntil Bool_Confirm=TRUE;
            WaitUntil Bool_Confirm=FALSE;
            MoveL Target_APuntosRef_110,Vel_Acercamiento,Z_Acercamiento,Prototipo_JSDaleman\WObj:=WO_PastelDef;
            WaitUntil Bool_Confirm=TRUE;
            WaitUntil Bool_Confirm=FALSE;
            MoveL Target_APuntosRef_120,Vel_Acercamiento,Z_Acercamiento,Prototipo_JSDaleman\WObj:=WO_PastelDef;
            MoveJ Target_APuntosRef_130,Vel_Vacio,Z_VacioMov,Prototipo_JSDaleman\WObj:=WO_PastelDef;
            WaitUntil Bool_Confirm=TRUE;
            WaitUntil Bool_Confirm=FALSE;
            MoveL Target_APuntosRef_140,Vel_Acercamiento,Z_Acercamiento,Prototipo_JSDaleman\WObj:=WO_PastelDef;
            WaitUntil Bool_Confirm=TRUE;
            WaitUntil Bool_Confirm=FALSE;
            MoveL Target_APuntosRef_150,Vel_Acercamiento,Z_Acercamiento,Prototipo_JSDaleman\WObj:=WO_PastelDef;
            MoveJ Target_RobLab_10,Vel_Vacio,Z_VacioMov,Prototipo_JSDaleman\WObj:=WO_PastelDef;
            WaitUntil Bool_Confirm=TRUE;
            WaitUntil Bool_Confirm=FALSE;
            MoveL Target_RobLab_20,Vel_Acercamiento,Z_Acercamiento,Prototipo_JSDaleman\WObj:=WO_PastelDef;
            WaitUntil Bool_Confirm=TRUE;
            WaitUntil Bool_Confirm=FALSE;
            MoveL Target_RobLab_260,Vel_Acercamiento,Z_Acercamiento,Prototipo_JSDaleman\WObj:=WO_PastelDef;
            WaitUntil Bool_Confirm=TRUE;
            WaitUntil Bool_Confirm=FALSE;
            MoveJ Target_Home_10,Vel_Vacio_Rap,Z_Vacio_Rap,Prototipo_JSDaleman\WObj:=wobj0;
            MoveJ Target_Frente_10,Vel_Vacio,Z_VacioMov,Prototipo_JSDaleman\WObj:=WO_PastelDef;
            MoveJ Target_Frente_20,Vel_Vacio,Z_VacioMov,Prototipo_JSDaleman\WObj:=WO_PastelDef;
            MoveJ Target_DibChip_10,Vel_Vacio,Z_VacioMov,Prototipo_JSDaleman\WObj:=WO_PastelDef;
            WaitUntil Bool_Confirm=TRUE;
            WaitUntil Bool_Confirm=FALSE;
            MoveL Target_DibChip_20,Vel_Proceso,Z_Proceso,Prototipo_JSDaleman\WObj:=WO_PastelDef;
            WaitUntil Bool_Confirm=TRUE;
            WaitUntil Bool_Confirm=FALSE;
            MoveL Target_DibChip_510,Vel_Acercamiento,Z_Acercamiento,Prototipo_JSDaleman\WObj:=WO_PastelDef;
            WaitUntil Bool_Confirm=TRUE;
            WaitUntil Bool_Confirm=FALSE;
            MoveJ Target_Frente_20,Vel_Vacio,Z_VacioMov,Prototipo_JSDaleman\WObj:=WO_PastelDef;
            MoveJ Target_Frente_10,Vel_Vacio,Z_VacioMov,Prototipo_JSDaleman\WObj:=WO_PastelDef;
            MoveJ Target_Home_10,Vel_Vacio_Rap,Z_Vacio_Rap,Prototipo_JSDaleman\WObj:=wobj0;
            MoveJ Target_Frente_30,Vel_Vacio_Rap,Z_Vacio_Rap,Prototipo_JSDaleman\WObj:=WO_PastelDef;
            MoveJ Target_Frente_40,Vel_Vacio_Rap,Z_Vacio_Rap,Prototipo_JSDaleman\WObj:=WO_PastelDef;
            MoveJ Target_DibEng_10,Vel_Vacio,Z_VacioMov,Prototipo_JSDaleman\WObj:=WO_PastelDef;
            WaitUntil Bool_Confirm=TRUE;
            WaitUntil Bool_Confirm=FALSE;
            MoveL Target_DibEng_20,Vel_Proceso,Z_Proceso,Prototipo_JSDaleman\WObj:=WO_PastelDef;
            WaitUntil Bool_Confirm=TRUE;
            WaitUntil Bool_Confirm=FALSE;
            MoveL Target_DibEng_790,Vel_Acercamiento,Z_Acercamiento,Prototipo_JSDaleman\WObj:=WO_PastelDef;
            WaitUntil Bool_Confirm=TRUE;
            WaitUntil Bool_Confirm=FALSE;
            MoveJ Target_Frente_40,Vel_Vacio_Rap,Z_Vacio_Rap,Prototipo_JSDaleman\WObj:=WO_PastelDef;
            MoveJ Target_Frente_30,Vel_Vacio_Rap,Z_Vacio_Rap,Prototipo_JSDaleman\WObj:=WO_PastelDef;
            MoveJ Target_Home_10,Vel_Vacio_Rap,Z_Paro,Prototipo_JSDaleman\WObj:=wobj0;
            Test_Transi:=TRUE;
        ENDIF
        RestoPath;
        StopMove;
        IEnable;
        CONNECT socket_com_in WITH SockDataIn;
        IPers cmd, socket_com_in;
    ENDTRAP
    TRAP Path_Parada
        IDelete socket_com_in;
        IDisable;
        StopMove;
        ClearPath;
        StorePath;
        Test_LabSIR:=FALSE;
        Test_25:=FALSE;
        Test_165:=FALSE;
        UIMsgBox \Header:="Parada ejecutada",
            mensaje_parada{1} \MsgLine2:=mensaje_parada{2} \MsgLine3:=mensaje_parada{3},
            \Buttons:=btnOK
            \Icon:=iconWarning
            \Result:=respuesta_parada;
        IWatch ReiniciarRut;
        WHILE Reiniciar <> TRUE DO
            Test_Reinicio:=TRUE;
            WaitTime 0.005;
            Test_Reinicio:=FALSE;
            WaitTime 0.005;
        ENDWHILE
        RestoPath;
        StopMove;
        IEnable;
        CONNECT socket_com_in WITH SockDataIn;
        IPers cmd, socket_com_in;
    ENDTRAP
    TRAP Path_PausCont
        IDelete socket_com_in;
        IDisable;
        ISleep PausaContinuar;
        StopMove;
        StorePath;
        WaitUntil Paus_Continue=TRUE;
        Paus_Continue:=FALSE;
        RestoPath;
        StartMove;
        WaitTime 0.1;
        IWatch PausaContinuar;
        IEnable;
        CONNECT socket_com_in WITH SockDataIn;
        IPers cmd, socket_com_in;
    ENDTRAP
    TRAP Path_Reinicio
        IDelete socket_com_in;
        IDisable;
        StopMove;
        ClearPath;
        StorePath;
        Test_LabSIR:=FALSE;
        Test_25:=FALSE;
        Test_165:=FALSE;
        Test_Reinicio:=TRUE;
        UIMsgBox \Header:="Reinicio ejecutado",
            mensaje_reinicio{1} \MsgLine2:=mensaje_reinicio{2} \MsgLine3:=mensaje_reinicio{3},
            \Buttons:=btnOK
            \Icon:=iconWarning
            \Result:=respuesta_parada;
        StartMove;
        MoveJ Target_Home_10,Vel_Vacio_Rap,Z_Vacio_Rap,Prototipo_JSDaleman\WObj:=wobj0;
        MoveJ Target_Espera,Vel_Vacio_Rap,Z_Paro,Prototipo_JSDaleman\WObj:=wobj0;
        Test_Reinicio:=FALSE;
        SetDO DO_03,1;
        RestoPath;
        StopMove;
        IEnable;
        ExitCycle;
    ENDTRAP
    TRAP IncIndicesContacto
        Incr index_contacto_origen;
        Incr index_contacto_destino;
    ENDTRAP
    TRAP IncIndicesContactoCir
        Incr index_contacto_origen;
        Incr index_contacto_origen;
        Incr index_contacto_destino;
        Incr index_contacto_destino;
    ENDTRAP
    TRAP IncIndicesVacio
        Incr index_vacio_origen;
    ENDTRAP
ENDMODULE

--- Controller Data/IRB140_LabSIR/RAPID/TASK1/PROGMOD/InterrupcionesSocket.mod ---
MODULE InterrupcionesSocket
    !***********************************************************
    !
    ! Modulo:  InterrupcionesSocket
    !
    ! Descripcion:
    !   Interrupciones generadas desde el socket
    !
    ! Autor: Juan_Daleman
    !
    ! Versión: 1.0
    !
    !***********************************************************

    !Variables de interrupcion
    VAR intnum SockParadaActiva;
    VAR intnum SockPausaActiva;
    VAR intnum SockBloqueoActiva;

    !Interrupción de lectura del socket
    VAR intnum socket_com_in;
    VAR intnum socket_com_out;

    !Variables de mensajes de error para el usuario
     VAR btnres respuesta_parada_socket;
     CONST string mensaje_parada_socket{3} := ["Parada del sistema ejecutada desde el socket", "Es necesario realizar rearme de operación", "Reinicie el sistema"];

    TRAP SockParada
        IDelete socket_com_in;
        IDisable;
        StopMove;
        ClearPath;
        StorePath;
        Sock_Parada:=FALSE;
        Test_LabSIR:=FALSE;
        Test_25:=FALSE;
        Test_165:=FALSE;
        UIMsgBox \Header:="Parada ejecutada",
            mensaje_parada_socket{1} \MsgLine2:=mensaje_parada_socket{2} \MsgLine3:=mensaje_parada_socket{3},
            \Buttons:=btnOK
            \Icon:=iconWarning
            \Result:=respuesta_parada;
        IWatch ReiniciarRut;
        WHILE Reiniciar <> TRUE DO
            Test_Reinicio:=TRUE;
            WaitTime 0.005;
            Test_Reinicio:=FALSE;
            WaitTime 0.005;
        ENDWHILE
        RestoPath;
        StopMove;
        IEnable;
        CONNECT socket_com_in WITH SockDataIn;
        IPers cmd, socket_com_in;
    ENDTRAP
    TRAP SockPausa
        IDelete socket_com_in;
        IDisable;
        ISleep PausaContinuar;
        ISleep SockPausaActiva;
        StopMove;
        StorePath;
        Sock_Pausa:=FALSE;
        WaitUntil Paus_Continue=TRUE;
        Paus_Continue:=FALSE;
        RestoPath;
        StartMove;
        WaitTime 0.1;
        IWatch PausaContinuar;
        IWatch SockPausaActiva;
        IEnable;
        CONNECT socket_com_in WITH SockDataIn;
        IPers cmd, socket_com_in;
    ENDTRAP
    TRAP SockBloqueo
        IDisable;
        ISleep SockBloqueoActiva;
        StopMove;
        IF NOT Postura_segura THEN
            StorePath;
            p_salida := CRobT(\Tool:=Prototipo_JSDaleman \WObj:=WO_PastelDef);
        ENDIF
        Sock_Bloquear:=FALSE;
        WHILE NOT Sock_Reinicio DO
            RevisarSocket;
        ENDWHILE
        Sock_Reinicio:=FALSE;
        RestoPath;
        Postura_segura:=FALSE;
        StartMove;
        WaitTime 0.1;
        IWatch SockBloqueoActiva;
        IEnable;
    ENDTRAP
    TRAP SockDataIn
        IDelete socket_com_in;
        IDisable;
        RevisarSocket;
        CONNECT socket_com_in WITH SockDataIn;
        IPers cmd, socket_com_in;
        IEnable;
    ENDTRAP
    TRAP SockDataOut
         WaitTime tiempo_envio;
    ENDTRAP
ENDMODULE

--- Controller Data/IRB140_LabSIR/RAPID/TASK1/PROGMOD/LABSIR.mod ---
MODULE LABSIR
    !***********************************************************
    !
    ! Modulo:  LABSIR
    !
    ! Descripción:
    !   Modulo con rutinas para decoracion con el motivo LABSIR
    !
    ! Autor: Juan_Daleman
    !
    ! Versión: 1.0
    !
    !***********************************************************

    !Puntos para diseno de la tapa
    !***********************************************************
    !Diseno de Robot de LabSir
    CONST robtarget Target_RobLab_10:=[[97.393,-56.932,-20],[0.707106781,0,0,0.707106781],[0,0,0,0],[9E+09,9E+09,9E+09,9E+09,9E+09,9E+09]];
    CONST robtarget Target_RobLab_20:=[[97.393,-56.932,0],[0.707106781,0,0,0.707106781],[0,0,0,0],[9E+09,9E+09,9E+09,9E+09,9E+09,9E+09]];
    CONST robtarget Target_RobLab_30:=[[27.685,-57.048,0],[0.707106781,0,0,0.707106781],[0,0,0,0],[9E+09,9E+09,9E+09,9E+09,9E+09,9E+09]];
    CONST robtarget Target_RobLab_40:=[[28.052,-51.495,0],[0.707106781,0,0,0.707106781],[0,0,0,0],[9E+09,9E+09,9E+09,9E+09,9E+09,9E+09]];
    CONST robtarget Target_RobLab_50:=[[30.377,-50.036,0],[0.707106781,0,0,0.707106781],[0,0,0,0],[9E+09,9E+09,9E+09,9E+09,9E+09,9E+09]];
    CONST robtarget Target_RobLab_60:=[[31.658,-49.677,0],[0.707106781,0,0,0.707106781],[0,0,0,0],[9E+09,9E+09,9E+09,9E+09,9E+09,9E+09]];
    CONST robtarget Target_RobLab_70:=[[32.366,-44.499,0],[0.707106781,0,0,0.707106781],[0,0,0,0],[9E+09,9E+09,9E+09,9E+09,9E+09,9E+09]];
    CONST robtarget Target_RobLab_80:=[[33.326,-43.358,0],[0.707106781,0,0,0.707106781],[0,0,0,0],[9E+09,9E+09,9E+09,9E+09,9E+09,9E+09]];
    CONST robtarget Target_RobLab_90:=[[35.236,-42.613,0],[0.707106781,0,0,0.707106781],[0,0,0,0],[9E+09,9E+09,9E+09,9E+09,9E+09,9E+09]];
    CONST robtarget Target_RobLab_100:=[[41.473,-42.079,0],[0.707106781,0,0,0.707106781],[0,0,0,0],[9E+09,9E+09,9E+09,9E+09,9E+09,9E+09]];
    CONST robtarget Target_RobLab_110:=[[42.167,-37.235,0],[0.707106781,0,0,0.707106781],[0,0,0,0],[9E+09,9E+09,9E+09,9E+09,9E+09,9E+09]];
    CONST robtarget Target_RobLab_120:=[[42.499,-36.72,0],[0.707106781,0,0,0.707106781],[0,0,0,0],[9E+09,9E+09,9E+09,9E+09,9E+09,9E+09]];
    CONST robtarget Target_RobLab_130:=[[42.787,-36.24,0],[0.707106781,0,0,0.707106781],[0,0,0,0],[9E+09,9E+09,9E+09,9E+09,9E+09,9E+09]];
    CONST robtarget Target_RobLab_140:=[[43.299,-35.809,0],[0.707106781,0,0,0.707106781],[0,0,0,0],[9E+09,9E+09,9E+09,9E+09,9E+09,9E+09]];
    CONST robtarget Target_RobLab_150:=[[45.768,-35.479,0],[0.707106781,0,0,0.707106781],[0,0,0,0],[9E+09,9E+09,9E+09,9E+09,9E+09,9E+09]];
    CONST robtarget Target_RobLab_160:=[[66.402,-35.529,0],[0.707106781,0,0,0.707106781],[0,0,0,0],[9E+09,9E+09,9E+09,9E+09,9E+09,9E+09]];
    CONST robtarget Target_RobLab_170:=[[69.206,-35.818,0],[0.707106781,0,0,0.707106781],[0,0,0,0],[9E+09,9E+09,9E+09,9E+09,9E+09,9E+09]];
    CONST robtarget Target_RobLab_180:=[[69.978,-36.514,0],[0.707106781,0,0,0.707106781],[0,0,0,0],[9E+09,9E+09,9E+09,9E+09,9E+09,9E+09]];
    CONST robtarget Target_RobLab_190:=[[70.361,-38.678,0],[0.707106781,0,0,0.707106781],[0,0,0,0],[9E+09,9E+09,9E+09,9E+09,9E+09,9E+09]];
    CONST robtarget Target_RobLab_200:=[[76.031,-38.349,0],[0.707106781,0,0,0.707106781],[0,0,0,0],[9E+09,9E+09,9E+09,9E+09,9E+09,9E+09]];
    CONST robtarget Target_RobLab_210:=[[92.824,-37.475,0],[0.707106781,0,0,0.707106781],[0,0,0,0],[9E+09,9E+09,9E+09,9E+09,9E+09,9E+09]];
    CONST robtarget Target_RobLab_220:=[[94.202,-38.373,0],[0.707106781,0,0,0.707106781],[0,0,0,0],[9E+09,9E+09,9E+09,9E+09,9E+09,9E+09]];
    CONST robtarget Target_RobLab_230:=[[95.549,-39.694,0],[0.707106781,0,0,0.707106781],[0,0,0,0],[9E+09,9E+09,9E+09,9E+09,9E+09,9E+09]];
    CONST robtarget Target_RobLab_240:=[[96.564,-41.561,0],[0.707106781,0,0,0.707106781],[0,0,0,0],[9E+09,9E+09,9E+09,9E+09,9E+09,9E+09]];
    CONST robtarget Target_RobLab_250:=[[97.393,-56.932,0],[0.707106781,0,0,0.707106781],[0,0,0,0],[9E+09,9E+09,9E+09,9E+09,9E+09,9E+09]];
    CONST robtarget Target_RobLab_260:=[[97.393003819,-56.932012397,-19.99997651],[0.707106781,0,0,0.707106781],[-1,0,-2,0],[9E+09,9E+09,9E+09,9E+09,9E+09,9E+09]];
    CONST robtarget Target_RobLab_270:=[[76.056,-31.592,-20],[0.707106781,0,0,0.707106781],[0,0,0,0],[9E+09,9E+09,9E+09,9E+09,9E+09,9E+09]];
    CONST robtarget Target_RobLab_280:=[[76.056,-31.592,0],[0.707106781,0,0,0.707106781],[0,0,0,0],[9E+09,9E+09,9E+09,9E+09,9E+09,9E+09]];
    CONST robtarget Target_RobLab_290:=[[73.184,-32.642,0],[0.707106781,0,0,0.707106781],[0,0,0,0],[9E+09,9E+09,9E+09,9E+09,9E+09,9E+09]];
    CONST robtarget Target_RobLab_300:=[[40.573,-32.639,0],[0.707106781,0,0,0.707106781],[0,0,0,0],[9E+09,9E+09,9E+09,9E+09,9E+09,9E+09]];
    CONST robtarget Target_RobLab_310:=[[38.777,-31.245,0],[0.707106781,0,0,0.707106781],[0,0,0,0],[9E+09,9E+09,9E+09,9E+09,9E+09,9E+09]];
    CONST robtarget Target_RobLab_320:=[[38.506,-29.103,0],[0.707106781,0,0,0.707106781],[0,0,0,0],[9E+09,9E+09,9E+09,9E+09,9E+09,9E+09]];
    CONST robtarget Target_RobLab_330:=[[30.583,-28.089,0],[0.707106781,0,0,0.707106781],[0,0,0,0],[9E+09,9E+09,9E+09,9E+09,9E+09,9E+09]];
    CONST robtarget Target_RobLab_340:=[[27.45,-26.522,0],[0.707106781,0,0,0.707106781],[0,0,0,0],[9E+09,9E+09,9E+09,9E+09,9E+09,9E+09]];
    CONST robtarget Target_RobLab_350:=[[25.478,-24.141,0],[0.707106781,0,0,0.707106781],[0,0,0,0],[9E+09,9E+09,9E+09,9E+09,9E+09,9E+09]];
    CONST robtarget Target_RobLab_360:=[[24.831,-22.791,0],[0.707106781,0,0,0.707106781],[0,0,0,0],[9E+09,9E+09,9E+09,9E+09,9E+09,9E+09]];
    CONST robtarget Target_RobLab_370:=[[24.858,-15.876,0],[0.707106781,0,0,0.707106781],[0,0,0,0],[9E+09,9E+09,9E+09,9E+09,9E+09,9E+09]];
    CONST robtarget Target_RobLab_380:=[[27.402,-4.781,0],[0.707106781,0,0,0.707106781],[0,0,0,0],[9E+09,9E+09,9E+09,9E+09,9E+09,9E+09]];
    CONST robtarget Target_RobLab_390:=[[28.59,-1.031,0],[0.707106781,0,0,0.707106781],[0,0,0,0],[9E+09,9E+09,9E+09,9E+09,9E+09,9E+09]];
    CONST robtarget Target_RobLab_400:=[[32.131,6.498,0],[0.707106781,0,0,0.707106781],[0,0,0,0],[9E+09,9E+09,9E+09,9E+09,9E+09,9E+09]];
    CONST robtarget Target_RobLab_410:=[[34.45,9.999,0],[0.707106781,0,0,0.707106781],[0,0,0,0],[9E+09,9E+09,9E+09,9E+09,9E+09,9E+09]];
    CONST robtarget Target_RobLab_420:=[[35.967,17.853,0],[0.707106781,0,0,0.707106781],[0,0,0,0],[9E+09,9E+09,9E+09,9E+09,9E+09,9E+09]];
    CONST robtarget Target_RobLab_430:=[[34.331,33.358,0],[0.707106781,0,0,0.707106781],[0,0,0,0],[9E+09,9E+09,9E+09,9E+09,9E+09,9E+09]];
    CONST robtarget Target_RobLab_440:=[[21.886,38.642,0],[0.707106781,0,0,0.707106781],[0,0,0,0],[9E+09,9E+09,9E+09,9E+09,9E+09,9E+09]];
    CONST robtarget Target_RobLab_450:=[[20.428,40.417,0],[0.707106781,0,0,0.707106781],[0,0,0,0],[9E+09,9E+09,9E+09,9E+09,9E+09,9E+09]];
    CONST robtarget Target_RobLab_460:=[[19.977,43.225,0],[0.707106781,0,0,0.707106781],[0,0,0,0],[9E+09,9E+09,9E+09,9E+09,9E+09,9E+09]];
    CONST robtarget Target_RobLab_470:=[[20.503,46.13,0],[0.707106781,0,0,0.707106781],[0,0,0,0],[9E+09,9E+09,9E+09,9E+09,9E+09,9E+09]];
    CONST robtarget Target_RobLab_480:=[[17.426,47.932,0],[0.707106781,0,0,0.707106781],[0,0,0,0],[9E+09,9E+09,9E+09,9E+09,9E+09,9E+09]];
    CONST robtarget Target_RobLab_490:=[[11.135,50.37,0],[0.707106781,0,0,0.707106781],[0,0,0,0],[9E+09,9E+09,9E+09,9E+09,9E+09,9E+09]];
    CONST robtarget Target_RobLab_500:=[[5.08,52.486,0],[0.707106781,0,0,0.707106781],[0,0,0,0],[9E+09,9E+09,9E+09,9E+09,9E+09,9E+09]];
    CONST robtarget Target_RobLab_510:=[[-5.504,56.417,0],[0.707106781,0,0,0.707106781],[0,0,0,0],[9E+09,9E+09,9E+09,9E+09,9E+09,9E+09]];
    CONST robtarget Target_RobLab_520:=[[-12.423,57.967,0],[0.707106781,0,0,0.707106781],[0,0,0,0],[9E+09,9E+09,9E+09,9E+09,9E+09,9E+09]];
    CONST robtarget Target_RobLab_530:=[[-14.489,58.698,0],[0.707106781,0,0,0.707106781],[0,0,0,0],[9E+09,9E+09,9E+09,9E+09,9E+09,9E+09]];
    CONST robtarget Target_RobLab_540:=[[-16.639,60.29,0],[0.707106781,0,0,0.707106781],[0,0,0,0],[9E+09,9E+09,9E+09,9E+09,9E+09,9E+09]];
    CONST robtarget Target_RobLab_550:=[[-18.331,62.54,0],[0.707106781,0,0,0.707106781],[0,0,0,0],[9E+09,9E+09,9E+09,9E+09,9E+09,9E+09]];
    CONST robtarget Target_RobLab_560:=[[-18.984,64.091,0],[0.707106781,0,0,0.707106781],[0,0,0,0],[9E+09,9E+09,9E+09,9E+09,9E+09,9E+09]];
    CONST robtarget Target_RobLab_570:=[[-19.206,66.036,0],[0.707106781,0,0,0.707106781],[0,0,0,0],[9E+09,9E+09,9E+09,9E+09,9E+09,9E+09]];
    CONST robtarget Target_RobLab_580:=[[-18.519,70.744,0],[0.707106781,0,0,0.707106781],[0,0,0,0],[9E+09,9E+09,9E+09,9E+09,9E+09,9E+09]];
    CONST robtarget Target_RobLab_590:=[[-15.337,74.49,0],[0.707106781,0,0,0.707106781],[0,0,0,0],[9E+09,9E+09,9E+09,9E+09,9E+09,9E+09]];
    CONST robtarget Target_RobLab_600:=[[-9.207,75.835,0],[0.707106781,0,0,0.707106781],[0,0,0,0],[9E+09,9E+09,9E+09,9E+09,9E+09,9E+09]];
    CONST robtarget Target_RobLab_610:=[[-6.76,75.294,0],[0.707106781,0,0,0.707106781],[0,0,0,0],[9E+09,9E+09,9E+09,9E+09,9E+09,9E+09]];
    CONST robtarget Target_RobLab_620:=[[-4.389,73.765,0],[0.707106781,0,0,0.707106781],[0,0,0,0],[9E+09,9E+09,9E+09,9E+09,9E+09,9E+09]];
    CONST robtarget Target_RobLab_630:=[[-2.968,72.434,0],[0.707106781,0,0,0.707106781],[0,0,0,0],[9E+09,9E+09,9E+09,9E+09,9E+09,9E+09]];
    CONST robtarget Target_RobLab_640:=[[1.54,70.372,0],[0.707106781,0,0,0.707106781],[0,0,0,0],[9E+09,9E+09,9E+09,9E+09,9E+09,9E+09]];
    CONST robtarget Target_RobLab_650:=[[5.693,71.178,0],[0.707106781,0,0,0.707106781],[0,0,0,0],[9E+09,9E+09,9E+09,9E+09,9E+09,9E+09]];
    CONST robtarget Target_RobLab_660:=[[16.189,67.574,0],[0.707106781,0,0,0.707106781],[0,0,0,0],[9E+09,9E+09,9E+09,9E+09,9E+09,9E+09]];
    CONST robtarget Target_RobLab_670:=[[17.8,66.343,0],[0.707106781,0,0,0.707106781],[0,0,0,0],[9E+09,9E+09,9E+09,9E+09,9E+09,9E+09]];
    CONST robtarget Target_RobLab_680:=[[19.62,63.596,0],[0.707106781,0,0,0.707106781],[0,0,0,0],[9E+09,9E+09,9E+09,9E+09,9E+09,9E+09]];
    CONST robtarget Target_RobLab_690:=[[24.48,61.692,0],[0.707106781,0,0,0.707106781],[0,0,0,0],[9E+09,9E+09,9E+09,9E+09,9E+09,9E+09]];
    CONST robtarget Target_RobLab_700:=[[27.685,63.964,0],[0.707106781,0,0,0.707106781],[0,0,0,0],[9E+09,9E+09,9E+09,9E+09,9E+09,9E+09]];
    CONST robtarget Target_RobLab_710:=[[30.828,64.206,0],[0.707106781,0,0,0.707106781],[0,0,0,0],[9E+09,9E+09,9E+09,9E+09,9E+09,9E+09]];
    CONST robtarget Target_RobLab_720:=[[32.382,63.772,0],[0.707106781,0,0,0.707106781],[0,0,0,0],[9E+09,9E+09,9E+09,9E+09,9E+09,9E+09]];
    CONST robtarget Target_RobLab_730:=[[35.068,64.958,0],[0.707106781,0,0,0.707106781],[0,0,0,0],[9E+09,9E+09,9E+09,9E+09,9E+09,9E+09]];
    CONST robtarget Target_RobLab_740:=[[37.198,65.238,0],[0.707106781,0,0,0.707106781],[0,0,0,0],[9E+09,9E+09,9E+09,9E+09,9E+09,9E+09]];
    CONST robtarget Target_RobLab_750:=[[42.544,63.627,0],[0.707106781,0,0,0.707106781],[0,0,0,0],[9E+09,9E+09,9E+09,9E+09,9E+09,9E+09]];
    CONST robtarget Target_RobLab_760:=[[57.898,57.969,0],[0.707106781,0,0,0.707106781],[0,0,0,0],[9E+09,9E+09,9E+09,9E+09,9E+09,9E+09]];
    CONST robtarget Target_RobLab_770:=[[65.982,52.123,0],[0.707106781,0,0,0.707106781],[0,0,0,0],[9E+09,9E+09,9E+09,9E+09,9E+09,9E+09]];
    CONST robtarget Target_RobLab_780:=[[65.262,38.5,0],[0.707106781,0,0,0.707106781],[0,0,0,0],[9E+09,9E+09,9E+09,9E+09,9E+09,9E+09]];
    CONST robtarget Target_RobLab_790:=[[63.087,33.606,0],[0.707106781,0,0,0.707106781],[0,0,0,0],[9E+09,9E+09,9E+09,9E+09,9E+09,9E+09]];
    CONST robtarget Target_RobLab_800:=[[60.923,30.286,0],[0.707106781,0,0,0.707106781],[0,0,0,0],[9E+09,9E+09,9E+09,9E+09,9E+09,9E+09]];
    CONST robtarget Target_RobLab_810:=[[57.281,27.367,0],[0.707106781,0,0,0.707106781],[0,0,0,0],[9E+09,9E+09,9E+09,9E+09,9E+09,9E+09]];
    CONST robtarget Target_RobLab_820:=[[57.475,18.633,0],[0.707106781,0,0,0.707106781],[0,0,0,0],[9E+09,9E+09,9E+09,9E+09,9E+09,9E+09]];
    CONST robtarget Target_RobLab_830:=[[55.509,8.537,0],[0.707106781,0,0,0.707106781],[0,0,0,0],[9E+09,9E+09,9E+09,9E+09,9E+09,9E+09]];
    CONST robtarget Target_RobLab_840:=[[58.351,1.091,0],[0.707106781,0,0,0.707106781],[0,0,0,0],[9E+09,9E+09,9E+09,9E+09,9E+09,9E+09]];
    CONST robtarget Target_RobLab_850:=[[58.469,-6.168,0],[0.707106781,0,0,0.707106781],[0,0,0,0],[9E+09,9E+09,9E+09,9E+09,9E+09,9E+09]];
    CONST robtarget Target_RobLab_860:=[[58.748,-13.963,0],[0.707106781,0,0,0.707106781],[0,0,0,0],[9E+09,9E+09,9E+09,9E+09,9E+09,9E+09]];
    CONST robtarget Target_RobLab_870:=[[63.065,-14.928,0],[0.707106781,0,0,0.707106781],[0,0,0,0],[9E+09,9E+09,9E+09,9E+09,9E+09,9E+09]];
    CONST robtarget Target_RobLab_880:=[[64.5,-17.412,0],[0.707106781,0,0,0.707106781],[0,0,0,0],[9E+09,9E+09,9E+09,9E+09,9E+09,9E+09]];
    CONST robtarget Target_RobLab_890:=[[66.248,-19.929,0],[0.707106781,0,0,0.707106781],[0,0,0,0],[9E+09,9E+09,9E+09,9E+09,9E+09,9E+09]];
    CONST robtarget Target_RobLab_900:=[[68.699,-20.675,0],[0.707106781,0,0,0.707106781],[0,0,0,0],[9E+09,9E+09,9E+09,9E+09,9E+09,9E+09]];
    CONST robtarget Target_RobLab_910:=[[71.718,-21.854,0],[0.707106781,0,0,0.707106781],[0,0,0,0],[9E+09,9E+09,9E+09,9E+09,9E+09,9E+09]];
    CONST robtarget Target_RobLab_920:=[[73.526,-22.54,0],[0.707106781,0,0,0.707106781],[0,0,0,0],[9E+09,9E+09,9E+09,9E+09,9E+09,9E+09]];
    CONST robtarget Target_RobLab_930:=[[75.108,-23.491,0],[0.707106781,0,0,0.707106781],[0,0,0,0],[9E+09,9E+09,9E+09,9E+09,9E+09,9E+09]];
    CONST robtarget Target_RobLab_940:=[[76.103,-25.055,0],[0.707106781,0,0,0.707106781],[0,0,0,0],[9E+09,9E+09,9E+09,9E+09,9E+09,9E+09]];
    CONST robtarget Target_RobLab_950:=[[76.056,-31.592,0],[0.707106781,0,0,0.707106781],[0,0,0,0],[9E+09,9E+09,9E+09,9E+09,9E+09,9E+09]];
    CONST robtarget Target_RobLab_960:=[[76.056,-31.592,-20],[0.707106781,0,0,0.707106781],[0,0,0,0],[9E+09,9E+09,9E+09,9E+09,9E+09,9E+09]];
    CONST robtarget Target_RobLab_970:=[[52.634,5.9,-20],[0.707106781,0,0,0.707106781],[0,0,0,0],[9E+09,9E+09,9E+09,9E+09,9E+09,9E+09]];
    CONST robtarget Target_RobLab_980:=[[52.634,5.9,0],[0.707106781,0,0,0.707106781],[0,0,0,0],[9E+09,9E+09,9E+09,9E+09,9E+09,9E+09]];
    CONST robtarget Target_RobLab_990:=[[50.793,7.747,0],[0.707106781,0,0,0.707106781],[0,0,0,0],[9E+09,9E+09,9E+09,9E+09,9E+09,9E+09]];
    CONST robtarget Target_RobLab_1000:=[[50.776,8.869,0],[0.707106781,0,0,0.707106781],[0,0,0,0],[9E+09,9E+09,9E+09,9E+09,9E+09,9E+09]];
    CONST robtarget Target_RobLab_1010:=[[51.246,10.934,0],[0.707106781,0,0,0.707106781],[0,0,0,0],[9E+09,9E+09,9E+09,9E+09,9E+09,9E+09]];
    CONST robtarget Target_RobLab_1020:=[[52.661,17.873,0],[0.707106781,0,0,0.707106781],[0,0,0,0],[9E+09,9E+09,9E+09,9E+09,9E+09,9E+09]];
    CONST robtarget Target_RobLab_1030:=[[52.746,24.375,0],[0.707106781,0,0,0.707106781],[0,0,0,0],[9E+09,9E+09,9E+09,9E+09,9E+09,9E+09]];
    CONST robtarget Target_RobLab_1040:=[[52.248,31.037,0],[0.707106781,0,0,0.707106781],[0,0,0,0],[9E+09,9E+09,9E+09,9E+09,9E+09,9E+09]];
    CONST robtarget Target_RobLab_1050:=[[52.178,32.951,0],[0.707106781,0,0,0.707106781],[0,0,0,0],[9E+09,9E+09,9E+09,9E+09,9E+09,9E+09]];
    CONST robtarget Target_RobLab_1060:=[[52.196,35.316,0],[0.707106781,0,0,0.707106781],[0,0,0,0],[9E+09,9E+09,9E+09,9E+09,9E+09,9E+09]];
    CONST robtarget Target_RobLab_1070:=[[52.671,36.092,0],[0.707106781,0,0,0.707106781],[0,0,0,0],[9E+09,9E+09,9E+09,9E+09,9E+09,9E+09]];
    CONST robtarget Target_RobLab_1080:=[[54.292,37.171,0],[0.707106781,0,0,0.707106781],[0,0,0,0],[9E+09,9E+09,9E+09,9E+09,9E+09,9E+09]];
    CONST robtarget Target_RobLab_1090:=[[54.614,33.296,0],[0.707106781,0,0,0.707106781],[0,0,0,0],[9E+09,9E+09,9E+09,9E+09,9E+09,9E+09]];
    CONST robtarget Target_RobLab_1100:=[[55.187,24.404,0],[0.707106781,0,0,0.707106781],[0,0,0,0],[9E+09,9E+09,9E+09,9E+09,9E+09,9E+09]];
    CONST robtarget Target_RobLab_1110:=[[55.197,18.369,0],[0.707106781,0,0,0.707106781],[0,0,0,0],[9E+09,9E+09,9E+09,9E+09,9E+09,9E+09]];
    CONST robtarget Target_RobLab_1120:=[[53.324,8.764,0],[0.707106781,0,0,0.707106781],[0,0,0,0],[9E+09,9E+09,9E+09,9E+09,9E+09,9E+09]];
    CONST robtarget Target_RobLab_1130:=[[52.634,5.9,0],[0.707106781,0,0,0.707106781],[0,0,0,0],[9E+09,9E+09,9E+09,9E+09,9E+09,9E+09]];
    CONST robtarget Target_RobLab_1140:=[[52.634,5.9,-20],[0.707106781,0,0,0.707106781],[0,0,0,0],[9E+09,9E+09,9E+09,9E+09,9E+09,9E+09]];
    CONST robtarget Target_RobLab_1150:=[[39.091,9.887,-20],[0.707106781,0,0,0.707106781],[0,0,0,0],[9E+09,9E+09,9E+09,9E+09,9E+09,9E+09]];
    CONST robtarget Target_RobLab_1160:=[[39.091,9.887,0],[0.707106781,0,0,0.707106781],[0,0,0,0],[9E+09,9E+09,9E+09,9E+09,9E+09,9E+09]];
    CONST robtarget Target_RobLab_1170:=[[36.875,8.762,0],[0.707106781,0,0,0.707106781],[0,0,0,0],[9E+09,9E+09,9E+09,9E+09,9E+09,9E+09]];
    CONST robtarget Target_RobLab_1180:=[[37.854,15.824,0],[0.707106781,0,0,0.707106781],[0,0,0,0],[9E+09,9E+09,9E+09,9E+09,9E+09,9E+09]];
    CONST robtarget Target_RobLab_1190:=[[38.057,18.938,0],[0.707106781,0,0,0.707106781],[0,0,0,0],[9E+09,9E+09,9E+09,9E+09,9E+09,9E+09]];
    CONST robtarget Target_RobLab_1200:=[[37.864,23.224,0],[0.707106781,0,0,0.707106781],[0,0,0,0],[9E+09,9E+09,9E+09,9E+09,9E+09,9E+09]];
    CONST robtarget Target_RobLab_1210:=[[37.429,28.804,0],[0.707106781,0,0,0.707106781],[0,0,0,0],[9E+09,9E+09,9E+09,9E+09,9E+09,9E+09]];
    CONST robtarget Target_RobLab_1220:=[[36.779,34.999,0],[0.707106781,0,0,0.707106781],[0,0,0,0],[9E+09,9E+09,9E+09,9E+09,9E+09,9E+09]];
    CONST robtarget Target_RobLab_1230:=[[38.457,34.571,0],[0.707106781,0,0,0.707106781],[0,0,0,0],[9E+09,9E+09,9E+09,9E+09,9E+09,9E+09]];
    CONST robtarget Target_RobLab_1240:=[[39.508,33.849,0],[0.707106781,0,0,0.707106781],[0,0,0,0],[9E+09,9E+09,9E+09,9E+09,9E+09,9E+09]];
    CONST robtarget Target_RobLab_1250:=[[40.153,28.462,0],[0.707106781,0,0,0.707106781],[0,0,0,0],[9E+09,9E+09,9E+09,9E+09,9E+09,9E+09]];
    CONST robtarget Target_RobLab_1260:=[[40.87,18.815,0],[0.707106781,0,0,0.707106781],[0,0,0,0],[9E+09,9E+09,9E+09,9E+09,9E+09,9E+09]];
    CONST robtarget Target_RobLab_1270:=[[39.908,13.523,0],[0.707106781,0,0,0.707106781],[0,0,0,0],[9E+09,9E+09,9E+09,9E+09,9E+09,9E+09]];
    CONST robtarget Target_RobLab_1280:=[[39.091,9.887,0],[0.707106781,0,0,0.707106781],[0,0,0,0],[9E+09,9E+09,9E+09,9E+09,9E+09,9E+09]];
    CONST robtarget Target_RobLab_1290:=[[39.091,9.887,-20],[0.707106781,0,0,0.707106781],[0,0,0,0],[9E+09,9E+09,9E+09,9E+09,9E+09,9E+09]];
    CONST robtarget Target_RobLab_1300:=[[45.877,-7.501,-20],[0.707106781,0,0,0.707106781],[0,0,0,0],[9E+09,9E+09,9E+09,9E+09,9E+09,9E+09]];
    CONST robtarget Target_RobLab_1310:=[[45.877,-7.501,0],[0.707106781,0,0,0.707106781],[0,0,0,0],[9E+09,9E+09,9E+09,9E+09,9E+09,9E+09]];
    CONST robtarget Target_RobLab_1320:=[[36.48,-0.258,0],[0.707106781,0,0,0.707106781],[0,0,0,0],[9E+09,9E+09,9E+09,9E+09,9E+09,9E+09]];
    CONST robtarget Target_RobLab_1330:=[[43.101,5.572,0],[0.707106781,0,0,0.707106781],[0,0,0,0],[9E+09,9E+09,9E+09,9E+09,9E+09,9E+09]];
    CONST robtarget Target_RobLab_1340:=[[50.085,-0.841,0],[0.707106781,0,0,0.707106781],[0,0,0,0],[9E+09,9E+09,9E+09,9E+09,9E+09,9E+09]];
    CONST robtarget Target_RobLab_1350:=[[45.877,-7.501,0],[0.707106781,0,0,0.707106781],[0,0,0,0],[9E+09,9E+09,9E+09,9E+09,9E+09,9E+09]];
    CONST robtarget Target_RobLab_1360:=[[45.877,-7.501,-20],[0.707106781,0,0,0.707106781],[0,0,0,0],[9E+09,9E+09,9E+09,9E+09,9E+09,9E+09]];
    CONST robtarget Target_RobLab_1370:=[[46.221,-10.037,-20],[0.707106781,0,0,0.707106781],[0,0,0,0],[9E+09,9E+09,9E+09,9E+09,9E+09,9E+09]];
    CONST robtarget Target_RobLab_1380:=[[46.221,-10.037,0],[0.707106781,0,0,0.707106781],[0,0,0,0],[9E+09,9E+09,9E+09,9E+09,9E+09,9E+09]];
    CONST robtarget Target_RobLab_1390:=[[33.996,-2.825,0],[0.707106781,0,0,0.707106781],[0,0,0,0],[9E+09,9E+09,9E+09,9E+09,9E+09,9E+09]];
    CONST robtarget Target_RobLab_1400:=[[40.131,7.626,0],[0.707106781,0,0,0.707106781],[0,0,0,0],[9E+09,9E+09,9E+09,9E+09,9E+09,9E+09]];
    CONST robtarget Target_RobLab_1410:=[[51.648,2.744,0],[0.707106781,0,0,0.707106781],[0,0,0,0],[9E+09,9E+09,9E+09,9E+09,9E+09,9E+09]];
    CONST robtarget Target_RobLab_1420:=[[46.221,-10.037,0],[0.707106781,0,0,0.707106781],[0,0,0,0],[9E+09,9E+09,9E+09,9E+09,9E+09,9E+09]];
    CONST robtarget Target_RobLab_1430:=[[46.221,-10.037,-20],[0.707106781,0,0,0.707106781],[0,0,0,0],[9E+09,9E+09,9E+09,9E+09,9E+09,9E+09]];
    CONST robtarget Target_RobLab_1440:=[[50.1,40.579,-20],[0.707106781,0,0,0.707106781],[0,0,0,0],[9E+09,9E+09,9E+09,9E+09,9E+09,9E+09]];
    CONST robtarget Target_RobLab_1450:=[[50.1,40.579,0],[0.707106781,0,0,0.707106781],[0,0,0,0],[9E+09,9E+09,9E+09,9E+09,9E+09,9E+09]];
    CONST robtarget Target_RobLab_1460:=[[36.843,43.426,0],[0.707106781,0,0,0.707106781],[0,0,0,0],[9E+09,9E+09,9E+09,9E+09,9E+09,9E+09]];
    CONST robtarget Target_RobLab_1470:=[[43.65824364,54.260056096,0],[0.707106781,0,0,0.707106781],[0,0,0,0],[9E+09,9E+09,9E+09,9E+09,9E+09,9E+09]];
    CONST robtarget Target_RobLab_1480:=[[50.491,51.546,0],[0.707106781,0,0,0.707106781],[0,0,0,0],[9E+09,9E+09,9E+09,9E+09,9E+09,9E+09]];
    CONST robtarget Target_RobLab_1490:=[[50.1,40.579,0],[0.707106781,0,0,0.707106781],[0,0,0,0],[9E+09,9E+09,9E+09,9E+09,9E+09,9E+09]];
    CONST robtarget Target_RobLab_1500:=[[50.1,40.579,-20],[0.707106781,0,0,0.707106781],[0,0,0,0],[9E+09,9E+09,9E+09,9E+09,9E+09,9E+09]];
    CONST robtarget Target_RobLab_1510:=[[47.789,35.991,-20],[0.707106781,0,0,0.707106781],[0,0,0,0],[9E+09,9E+09,9E+09,9E+09,9E+09,9E+09]];
    CONST robtarget Target_RobLab_1520:=[[47.789,35.991,0],[0.707106781,0,0,0.707106781],[0,0,0,0],[9E+09,9E+09,9E+09,9E+09,9E+09,9E+09]];
    CONST robtarget Target_RobLab_1530:=[[33.611,46.793,0],[0.707106781,0,0,0.707106781],[0,0,0,0],[9E+09,9E+09,9E+09,9E+09,9E+09,9E+09]];
    CONST robtarget Target_RobLab_1540:=[[46.858,56.902,0],[0.707106781,0,0,0.707106781],[0,0,0,0],[9E+09,9E+09,9E+09,9E+09,9E+09,9E+09]];
    CONST robtarget Target_RobLab_1550:=[[55.247,46.149,0],[0.707106781,0,0,0.707106781],[0,0,0,0],[9E+09,9E+09,9E+09,9E+09,9E+09,9E+09]];
    CONST robtarget Target_RobLab_1560:=[[47.789,35.991,0],[0.707106781,0,0,0.707106781],[0,0,0,0],[9E+09,9E+09,9E+09,9E+09,9E+09,9E+09]];
    CONST robtarget Target_RobLab_1570:=[[47.789,35.991,-20],[0.707106781,0,0,0.707106781],[0,0,0,0],[9E+09,9E+09,9E+09,9E+09,9E+09,9E+09]];
    CONST robtarget Target_RobLab_1580:=[[-6.147,64.723,-20],[0.707106781,0,0,0.707106781],[0,0,0,0],[9E+09,9E+09,9E+09,9E+09,9E+09,9E+09]];
    CONST robtarget Target_RobLab_1590:=[[-6.147,64.723,0],[0.707106781,0,0,0.707106781],[0,0,0,0],[9E+09,9E+09,9E+09,9E+09,9E+09,9E+09]];
    CONST robtarget Target_RobLab_1600:=[[-13.254,63.189,0],[0.707106781,0,0,0.707106781],[0,0,0,0],[9E+09,9E+09,9E+09,9E+09,9E+09,9E+09]];
    CONST robtarget Target_RobLab_1610:=[[-12.004,71.159,0],[0.707106781,0,0,0.707106781],[0,0,0,0],[9E+09,9E+09,9E+09,9E+09,9E+09,9E+09]];
    CONST robtarget Target_RobLab_1620:=[[-6.512,69.605,0],[0.707106781,0,0,0.707106781],[0,0,0,0],[9E+09,9E+09,9E+09,9E+09,9E+09,9E+09]];
    CONST robtarget Target_RobLab_1630:=[[-5.611,66.562,0],[0.707106781,0,0,0.707106781],[0,0,0,0],[9E+09,9E+09,9E+09,9E+09,9E+09,9E+09]];
    CONST robtarget Target_RobLab_1640:=[[-6.147,64.723,-20],[0.707106781,0,0,0.707106781],[0,0,0,0],[9E+09,9E+09,9E+09,9E+09,9E+09,9E+09]];
    CONST robtarget Target_RobLab_1650:=[[-7.452,60.521,-20],[0.707106781,0,0,0.707106781],[0,0,0,0],[9E+09,9E+09,9E+09,9E+09,9E+09,9E+09]];
    CONST robtarget Target_RobLab_1660:=[[-7.452,60.521,0],[0.707106781,0,0,0.707106781],[0,0,0,0],[9E+09,9E+09,9E+09,9E+09,9E+09,9E+09]];
    CONST robtarget Target_RobLab_1670:=[[-16.57,64.05,0],[0.707106781,0,0,0.707106781],[0,0,0,0],[9E+09,9E+09,9E+09,9E+09,9E+09,9E+09]];
    CONST robtarget Target_RobLab_1680:=[[-12.72,73.276,0],[0.707106781,0,0,0.707106781],[0,0,0,0],[9E+09,9E+09,9E+09,9E+09,9E+09,9E+09]];
    CONST robtarget Target_RobLab_1690:=[[-3.568,65.694,0],[0.707106781,0,0,0.707106781],[0,0,0,0],[9E+09,9E+09,9E+09,9E+09,9E+09,9E+09]];
    CONST robtarget Target_RobLab_1700:=[[-7.452,60.521,0],[0.707106781,0,0,0.707106781],[0,0,0,0],[9E+09,9E+09,9E+09,9E+09,9E+09,9E+09]];
    CONST robtarget Target_RobLab_1710:=[[-7.452,60.521,-20],[0.707106781,0,0,0.707106781],[0,0,0,0],[9E+09,9E+09,9E+09,9E+09,9E+09,9E+09]];
    !**********************************************************
    !Dise?o de nombre LabSir
    CONST robtarget Target_10NomLab_L:=[[3.79755,47.324448,-20],[0.707106781,0,0,0.707106781],[0,0,0,0],[9E+09,9E+09,9E+09,9E+09,9E+09,9E+09]];
    CONST robtarget Target_20NomLab_L:=[[3.79755,47.324448,0],[0.707106781,0,0,0.707106781],[0,0,0,0],[9E+09,9E+09,9E+09,9E+09,9E+09,9E+09]];
    CONST robtarget Target_30NomLab_L:=[[2.597069625,3.348416,0],[0.707106781,0,0,0.707106781],[0,0,0,0],[9E+09,9E+09,9E+09,9E+09,9E+09,9E+09]];
    CONST robtarget Target_40NomLab_L:=[[-1.998180875,0.1710675,0],[0.707106781,0,0,0.707106781],[0,0,0,0],[9E+09,9E+09,9E+09,9E+09,9E+09,9E+09]];
    CONST robtarget Target_50NomLab_L:=[[-9.708635,-0.116667,0],[0.707106781,0,0,0.707106781],[0,0,0,0],[9E+09,9E+09,9E+09,9E+09,9E+09,9E+09]];
    CONST robtarget Target_60NomLab_L:=[[-9.708635,5.12076,0],[0.707106781,0,0,0.707106781],[0,0,0,0],[9E+09,9E+09,9E+09,9E+09,9E+09,9E+09]];
    CONST robtarget Target_70NomLab_L:=[[-1.286154,6.56909,0],[0.707106781,0,0,0.707106781],[0,0,0,0],[9E+09,9E+09,9E+09,9E+09,9E+09,9E+09]];
    CONST robtarget Target_80NomLab_L:=[[-1.286154,47.476319,0],[0.707106781,0,0,0.707106781],[0,0,0,0],[9E+09,9E+09,9E+09,9E+09,9E+09,9E+09]];
    CONST robtarget Target_90NomLab_L:=[[3.79755,47.324448,0],[0.707106781,0,0,0.707106781],[0,0,0,0],[9E+09,9E+09,9E+09,9E+09,9E+09,9E+09]];
    CONST robtarget Target_10NomLab_A:=[[-44.486792,29.956669,-20],[0.707106781,0,0,0.707106781],[0,0,0,0],[9E+09,9E+09,9E+09,9E+09,9E+09,9E+09]];
    CONST robtarget Target_20NomLab_A:=[[-44.486792,29.956669,0],[0.707106781,0,0,0.707106781],[0,0,0,0],[9E+09,9E+09,9E+09,9E+09,9E+09,9E+09]];
    CONST robtarget Target_30NomLab_A:=[[-45.446965,20.377958,0],[0.707106781,0,0,0.707106781],[0,-1,0,0],[9E+09,9E+09,9E+09,9E+09,9E+09,9E+09]];
    CONST robtarget Target_40NomLab_A:=[[-14.033515,20.377958,0],[0.707106781,0,0,0.707106781],[0,-1,0,0],[9E+09,9E+09,9E+09,9E+09,9E+09,9E+09]];
    CONST robtarget Target_50NomLab_A:=[[-14.912725,3.965854,0],[0.707106781,0,0,0.707106781],[0,-1,0,0],[9E+09,9E+09,9E+09,9E+09,9E+09,9E+09]];
    CONST robtarget Target_60NomLab_A:=[[-19.425723,0.264069,0],[0.707106781,0,0,0.707106781],[0,-1,0,0],[9E+09,9E+09,9E+09,9E+09,9E+09,9E+09]];
    CONST robtarget Target_70NomLab_A:=[[-50.454998,-0.116667,0],[0.707106781,0,0,0.707106781],[0,-1,0,0],[9E+09,9E+09,9E+09,9E+09,9E+09,9E+09]];
    CONST robtarget Target_80NomLab_A:=[[-49.995417,30.69565,0],[0.707106781,0,0,0.707106781],[0,-1,0,0],[9E+09,9E+09,9E+09,9E+09,9E+09,9E+09]];
    CONST robtarget Target_90NomLab_A:=[[-45.087396,35.436719,0],[0.707106781,0,0,0.707106781],[0,-1,0,0],[9E+09,9E+09,9E+09,9E+09,9E+09,9E+09]];
    CONST robtarget Target_100NomLab_A:=[[-14.033515,35.635156,0],[0.707106781,0,0,0.707106781],[0,-1,0,0],[9E+09,9E+09,9E+09,9E+09,9E+09,9E+09]];
    CONST robtarget Target_110NomLab_A:=[[-14.033515,30.625271,0],[0.707106781,0,0,0.707106781],[0,-1,0,0],[9E+09,9E+09,9E+09,9E+09,9E+09,9E+09]];
    CONST robtarget Target_120NomLab_A:=[[-44.486792,29.956669,0],[0.707106781,0,0,0.707106781],[0,-1,0,0],[9E+09,9E+09,9E+09,9E+09,9E+09,9E+09]];
    CONST robtarget Target_10NomLab_Aint:=[[-45.191377,15.060362,-20],[0.707106781,0,0,0.707106781],[0,0,0,0],[9E+09,9E+09,9E+09,9E+09,9E+09,9E+09]];
    CONST robtarget Target_20NomLab_Aint:=[[-45.191377,15.060362,0],[0.707106781,0,0,0.707106781],[0,0,0,0],[9E+09,9E+09,9E+09,9E+09,9E+09,9E+09]];
    CONST robtarget Target_30NomLab_Aint:=[[-45.333194,5.234796,0],[0.707106781,0,0,0.707106781],[0,0,0,0],[9E+09,9E+09,9E+09,9E+09,9E+09,9E+09]];
    CONST robtarget Target_40NomLab_Aint:=[[-20.275035,5.361796,0],[0.707106781,0,0,0.707106781],[0,0,0,0],[9E+09,9E+09,9E+09,9E+09,9E+09,9E+09]];
    CONST robtarget Target_50NomLab_Aint:=[[-19.041548,15.342144,0],[0.707106781,0,0,0.707106781],[0,0,0,0],[9E+09,9E+09,9E+09,9E+09,9E+09,9E+09]];
    CONST robtarget Target_60NomLab_Aint:=[[-45.191377,15.060362,0],[0.707106781,0,0,0.707106781],[0,0,0,0],[9E+09,9E+09,9E+09,9E+09,9E+09,9E+09]];
    CONST robtarget Target_10NomLab_B:=[[-70.800398,-0.116667,-20],[0.707106781,0,0,0.707106781],[0,-1,0,0],[9E+09,9E+09,9E+09,9E+09,9E+09,9E+09]];
    CONST robtarget Target_20NomLab_B:=[[-70.800398,-0.116667,0],[0.707106781,0,0,0.707106781],[0,0,0,0],[9E+09,9E+09,9E+09,9E+09,9E+09,9E+09]];
    CONST robtarget Target_30NomLab_B:=[[-88.365821,0.91071,0],[0.707106781,0,0,0.707106781],[0,0,0,0],[9E+09,9E+09,9E+09,9E+09,9E+09,9E+09]];
    CONST robtarget Target_40NomLab_B:=[[-92.0476305,7.729816625,0],[0.707106781,0,0,0.707106781],[0,0,0,0],[9E+09,9E+09,9E+09,9E+09,9E+09,9E+09]];
    CONST robtarget Target_50NomLab_B:=[[-90.973554,32.296115,0],[0.707106781,0,0,0.707106781],[0,0,0,0],[9E+09,9E+09,9E+09,9E+09,9E+09,9E+09]];
    CONST robtarget Target_60NomLab_B:=[[-87.050048,35.424019,0],[0.707106781,0,0,0.707106781],[0,0,0,0],[9E+09,9E+09,9E+09,9E+09,9E+09,9E+09]];
    CONST robtarget Target_70NomLab_B:=[[-60.760221375,36.8803515,0],[0.707106781,0,0,0.707106781],[0,0,0,0],[9E+09,9E+09,9E+09,9E+09,9E+09,9E+09]];
    CONST robtarget Target_80NomLab_B:=[[-60.698342,47.476319,0],[0.707106781,0,0,0.707106781],[0,0,0,0],[9E+09,9E+09,9E+09,9E+09,9E+09,9E+09]];
    CONST robtarget Target_90NomLab_B:=[[-55.690573,47.476319,0],[0.707106781,0,0,0.707106781],[0,0,0,0],[9E+09,9E+09,9E+09,9E+09,9E+09,9E+09]];
    CONST robtarget Target_100NomLab_B:=[[-55.690573,-0.116667,0],[0.707106781,0,0,0.707106781],[0,0,0,0],[9E+09,9E+09,9E+09,9E+09,9E+09,9E+09]];
    CONST robtarget Target_110NomLab_B:=[[-70.800398,-0.116667,0],[0.707106781,0,0,0.707106781],[0,0,0,0],[9E+09,9E+09,9E+09,9E+09,9E+09,9E+09]];
    CONST robtarget Target_10NomLab_Bint:=[[-86.202058,29.967252,-20],[0.707106781,0,0,0.707106781],[0,0,0,0],[9E+09,9E+09,9E+09,9E+09,9E+09,9E+09]];
    CONST robtarget Target_20NomLab_Bint:=[[-86.202058,29.967252,0],[0.707106781,0,0,0.707106781],[0,0,0,0],[9E+09,9E+09,9E+09,9E+09,9E+09,9E+09]];
    CONST robtarget Target_30NomLab_Bint:=[[-86.321385,5.818996,0],[0.707106781,0,0,0.707106781],[0,0,0,0],[9E+09,9E+09,9E+09,9E+09,9E+09,9E+09]];
    CONST robtarget Target_40NomLab_Bint:=[[-61.534425,5.843338,0],[0.707106781,0,0,0.707106781],[0,0,0,0],[9E+09,9E+09,9E+09,9E+09,9E+09,9E+09]];
    CONST robtarget Target_50NomLab_Bint:=[[-61.592898,29.928094,0],[0.707106781,0,0,0.707106781],[0,0,0,0],[9E+09,9E+09,9E+09,9E+09,9E+09,9E+09]];
    CONST robtarget Target_60NomLab_Bint:=[[-86.202058,29.967252,0],[0.707106781,0,0,0.707106781],[0,0,0,0],[9E+09,9E+09,9E+09,9E+09,9E+09,9E+09]];
    CONST robtarget Target_10NomLab_S:=[[3.133975,-12.610292,-20],[0.707106781,0,0,0.707106781],[0,0,0,0],[9E+09,9E+09,9E+09,9E+09,9E+09,9E+09]];
    CONST robtarget Target_20NomLab_S:=[[3.133975,-12.610292,0],[0.707106781,0,0,0.707106781],[0,0,0,0],[9E+09,9E+09,9E+09,9E+09,9E+09,9E+09]];
    CONST robtarget Target_30NomLab_S:=[[10.437004,-18.903406,0],[0.707106781,0,0,0.707106781],[0,0,0,0],[9E+09,9E+09,9E+09,9E+09,9E+09,9E+09]];
    CONST robtarget Target_40NomLab_S:=[[9.772106,-34.450058,0],[0.707106781,0,0,0.707106781],[0,0,0,0],[9E+09,9E+09,9E+09,9E+09,9E+09,9E+09]];
    CONST robtarget Target_50NomLab_S:=[[4.860117,-38.959088,0],[0.707106781,0,0,0.707106781],[0,0,0,0],[9E+09,9E+09,9E+09,9E+09,9E+09,9E+09]];
    CONST robtarget Target_60NomLab_S:=[[-23.935546,-39.625838,0],[0.707106781,0,0,0.707106781],[0,0,0,0],[9E+09,9E+09,9E+09,9E+09,9E+09,9E+09]];
    CONST robtarget Target_70NomLab_S:=[[-23.935546,-47.140533,0],[0.707106781,0,0,0.707106781],[0,0,0,0],[9E+09,9E+09,9E+09,9E+09,9E+09,9E+09]];
    CONST robtarget Target_80NomLab_S:=[[0.973917,-47.368075,0],[0.707106781,0,0,0.707106781],[0,0,0,0],[9E+09,9E+09,9E+09,9E+09,9E+09,9E+09]];
    CONST robtarget Target_90NomLab_S:=[[1.104092,-43.724763,0],[0.707106781,0,0,0.707106781],[0,0,0,0],[9E+09,9E+09,9E+09,9E+09,9E+09,9E+09]];
    CONST robtarget Target_100NomLab_S:=[[10.550775,-43.601467,0],[0.707106781,0,0,0.707106781],[0,0,0,0],[9E+09,9E+09,9E+09,9E+09,9E+09,9E+09]];
    CONST robtarget Target_110NomLab_S:=[[8.714037,-53.402692,0],[0.707106781,0,0,0.707106781],[0,0,0,0],[9E+09,9E+09,9E+09,9E+09,9E+09,9E+09]];
    CONST robtarget Target_120NomLab_S:=[[2.923631,-56.786713,0],[0.707106781,0,0,0.707106781],[0,0,0,0],[9E+09,9E+09,9E+09,9E+09,9E+09,9E+09]];
    CONST robtarget Target_130NomLab_S:=[[-26.667104,-56.674,0],[0.707106781,0,0,0.707106781],[0,0,0,0],[9E+09,9E+09,9E+09,9E+09,9E+09,9E+09]];
    CONST robtarget Target_140NomLab_S:=[[-32.793233875,-51.677079125,0],[0.707106781,0,0,0.707106781],[0,0,0,0],[9E+09,9E+09,9E+09,9E+09,9E+09,9E+09]];
    CONST robtarget Target_150NomLab_S:=[[-32.840263125,-35.198696625,0],[0.707106781,0,0,0.707106781],[0,0,0,0],[9E+09,9E+09,9E+09,9E+09,9E+09,9E+09]];
    CONST robtarget Target_160NomLab_S:=[[-26.023637,-29.974631,0],[0.707106781,0,0,0.707106781],[0,0,0,0],[9E+09,9E+09,9E+09,9E+09,9E+09,9E+09]];
    CONST robtarget Target_170NomLab_S:=[[0.990321,-29.720102,0],[0.707106781,0,0,0.707106781],[0,0,0,0],[9E+09,9E+09,9E+09,9E+09,9E+09,9E+09]];
    CONST robtarget Target_180NomLab_S:=[[0.990585,-22.091371,0],[0.707106781,0,0,0.707106781],[0,0,0,0],[9E+09,9E+09,9E+09,9E+09,9E+09,9E+09]];
    CONST robtarget Target_190NomLab_S:=[[-23.979532875,-22.814046875,0],[0.707106781,0,0,0.707106781],[0,0,0,0],[9E+09,9E+09,9E+09,9E+09,9E+09,9E+09]];
    CONST robtarget Target_200NomLab_S:=[[-24.049317,-25.848719,0],[0.707106781,0,0,0.707106781],[0,0,0,0],[9E+09,9E+09,9E+09,9E+09,9E+09,9E+09]];
    CONST robtarget Target_210NomLab_S:=[[-33.837577,-25.848719,0],[0.707106781,0,0,0.707106781],[0,0,0,0],[9E+09,9E+09,9E+09,9E+09,9E+09,9E+09]];
    CONST robtarget Target_220NomLab_S:=[[-31.20606425,-15.42115925,0],[0.707106781,0,0,0.707106781],[0,0,0,0],[9E+09,9E+09,9E+09,9E+09,9E+09,9E+09]];
    CONST robtarget Target_230NomLab_S:=[[-25.843456,-12.413442,0],[0.707106781,0,0,0.707106781],[0,0,0,0],[9E+09,9E+09,9E+09,9E+09,9E+09,9E+09]];
    CONST robtarget Target_240NomLab_S:=[[3.133975,-12.610292,0],[0.707106781,0,0,0.707106781],[0,0,0,0],[9E+09,9E+09,9E+09,9E+09,9E+09,9E+09]];
    CONST robtarget Target_05NomLab_I:=[[-39.178192,-12.698133,-20],[0.707106781,0,0,0.707106781],[0,0,0,0],[9E+09,9E+09,9E+09,9E+09,9E+09,9E+09]];
    CONST robtarget Target_10NomLab_I:=[[-39.178192,-12.698133,-20],[0.707106781,0,0,0.707106781],[0,0,0,0],[9E+09,9E+09,9E+09,9E+09,9E+09,9E+09]];
    CONST robtarget Target_20NomLab_I:=[[-39.178192,-12.698133,0],[0.707106781,0,0,0.707106781],[0,0,0,0],[9E+09,9E+09,9E+09,9E+09,9E+09,9E+09]];
    CONST robtarget Target_30NomLab_I:=[[-39.186923,-56.932233,0],[0.707106781,0,0,0.707106781],[0,0,0,0],[9E+09,9E+09,9E+09,9E+09,9E+09,9E+09]];
    CONST robtarget Target_40NomLab_I:=[[-48.633871,-57.055529,0],[0.707106781,0,0,0.707106781],[0,0,0,0],[9E+09,9E+09,9E+09,9E+09,9E+09,9E+09]];
    CONST robtarget Target_50NomLab_I:=[[-48.633871,-12.413442,0],[0.707106781,0,0,0.707106781],[0,0,0,0],[9E+09,9E+09,9E+09,9E+09,9E+09,9E+09]];
    CONST robtarget Target_60NomLab_I:=[[-39.178192,-12.698133,0],[0.707106781,0,0,0.707106781],[0,0,0,0],[9E+09,9E+09,9E+09,9E+09,9E+09,9E+09]];
    CONST robtarget Target_05NomLab_R:=[[-53.243442,-12.562931,-20],[0.707106781,0,0,0.707106781],[0,0,0,0],[9E+09,9E+09,9E+09,9E+09,9E+09,9E+09]];
    CONST robtarget Target_10NomLab_R:=[[-53.243442,-12.562931,-20],[0.707106781,0,0,0.707106781],[0,0,0,0],[9E+09,9E+09,9E+09,9E+09,9E+09,9E+09]];
    CONST robtarget Target_20NomLab_R:=[[-53.243442,-12.562931,0],[0.707106781,0,0,0.707106781],[0,0,0,0],[9E+09,9E+09,9E+09,9E+09,9E+09,9E+09]];
    CONST robtarget Target_30NomLab_R:=[[-52.95875,-57.055529,0],[0.707106781,0,0,0.707106781],[0,0,0,0],[9E+09,9E+09,9E+09,9E+09,9E+09,9E+09]];
    CONST robtarget Target_40NomLab_R:=[[-62.405698,-56.932233,0],[0.707106781,0,0,0.707106781],[0,0,0,0],[9E+09,9E+09,9E+09,9E+09,9E+09,9E+09]];
    CONST robtarget Target_50NomLab_R:=[[-62.525819,-42.543663,0],[0.707106781,0,0,0.707106781],[0,0,0,0],[9E+09,9E+09,9E+09,9E+09,9E+09,9E+09]];
    CONST robtarget Target_60NomLab_R:=[[-76.007133,-43.470763,0],[0.707106781,0,0,0.707106781],[0,0,0,0],[9E+09,9E+09,9E+09,9E+09,9E+09,9E+09]];
    CONST robtarget Target_70NomLab_R:=[[-87.563869,-57.055265,0],[0.707106781,0,0,0.707106781],[0,0,0,0],[9E+09,9E+09,9E+09,9E+09,9E+09,9E+09]];
    CONST robtarget Target_80NomLab_R:=[[-97.233596,-56.932233,0],[0.707106781,0,0,0.707106781],[0,0,0,0],[9E+09,9E+09,9E+09,9E+09,9E+09,9E+09]];
    CONST robtarget Target_90NomLab_R:=[[-95.014006,-50.87645,0],[0.707106781,0,0,0.707106781],[0,0,0,0],[9E+09,9E+09,9E+09,9E+09,9E+09,9E+09]];
    CONST robtarget Target_100NomLab_R:=[[-88.582646625,-42.2683965,0],[0.707106781,0,0,0.707106781],[0,0,0,0],[9E+09,9E+09,9E+09,9E+09,9E+09,9E+09]];
    CONST robtarget Target_110NomLab_R:=[[-96.168912,-37.385346,0],[0.707106781,0,0,0.707106781],[0,0,0,0],[9E+09,9E+09,9E+09,9E+09,9E+09,9E+09]];
    CONST robtarget Target_120NomLab_R:=[[-96.036725312,-17.219842617,0],[0.707106781,0,0,0.707106781],[0,0,0,0],[9E+09,9E+09,9E+09,9E+09,9E+09,9E+09]];
    CONST robtarget Target_130NomLab_R:=[[-91.922615,-13.372292,0],[0.707106781,0,0,0.707106781],[0,0,0,0],[9E+09,9E+09,9E+09,9E+09,9E+09,9E+09]];
    CONST robtarget Target_140NomLab_R:=[[-53.243442,-12.562931,0],[0.707106781,0,0,0.707106781],[0,0,0,0],[9E+09,9E+09,9E+09,9E+09,9E+09,9E+09]];
    CONST robtarget Target_05NomLab_Rint:=[[-87.50619,-27.43225,-20],[0.707106781,0,0,0.707106781],[0,0,0,0],[9E+09,9E+09,9E+09,9E+09,9E+09,9E+09]];
    CONST robtarget Target_10NomLab_Rint:=[[-87.50619,-27.43225,-20],[0.707106781,0,0,0.707106781],[0,0,0,0],[9E+09,9E+09,9E+09,9E+09,9E+09,9E+09]];
    CONST robtarget Target_20NomLab_Rint:=[[-87.50619,-27.43225,0],[0.707106781,0,0,0.707106781],[0,0,0,0],[9E+09,9E+09,9E+09,9E+09,9E+09,9E+09]];
    CONST robtarget Target_30NomLab_Rint:=[[-87.567573,-32.68026,0],[0.707106781,0,0,0.707106781],[0,0,0,0],[9E+09,9E+09,9E+09,9E+09,9E+09,9E+09]];
    CONST robtarget Target_40NomLab_Rint:=[[-62.519469,-32.68026,0],[0.707106781,0,0,0.707106781],[0,0,0,0],[9E+09,9E+09,9E+09,9E+09,9E+09,9E+09]];
    CONST robtarget Target_50NomLab_Rint:=[[-62.519469,-22.091371,0],[0.707106781,0,0,0.707106781],[0,0,0,0],[9E+09,9E+09,9E+09,9E+09,9E+09,9E+09]];
    CONST robtarget Target_60NomLab_Rint:=[[-87.445335,-22.18424,0],[0.707106781,0,0,0.707106781],[0,0,0,0],[9E+09,9E+09,9E+09,9E+09,9E+09,9E+09]];
    CONST robtarget Target_70NomLab_Rint:=[[-87.50619,-27.43225,0],[0.707106781,0,0,0.707106781],[0,0,0,0],[9E+09,9E+09,9E+09,9E+09,9E+09,9E+09]];
    CONST robtarget Target_100NomLab_L:=[[3.79755,47.324448,-20],[0.707106781,0,0,0.707106781],[0,0,0,0],[9E+09,9E+09,9E+09,9E+09,9E+09,9E+09]];
    CONST robtarget Target_130NomLab_A:=[[-44.486792,29.956669,-20],[0.707106781,0,0,0.707106781],[0,-1,0,0],[9E+09,9E+09,9E+09,9E+09,9E+09,9E+09]];
    CONST robtarget Target_70NomLab_Aint:=[[-45.191377,15.060362,-20],[0.707106781,0,0,0.707106781],[0,0,0,0],[9E+09,9E+09,9E+09,9E+09,9E+09,9E+09]];
    CONST robtarget Target_70NomLab_Bint:=[[-86.202058,29.967252,-20],[0.707106781,0,0,0.707106781],[0,0,0,0],[9E+09,9E+09,9E+09,9E+09,9E+09,9E+09]];
    CONST robtarget Target_250NomLab_S:=[[3.133975,-12.610292,-20],[0.707106781,0,0,0.707106781],[0,0,0,0],[9E+09,9E+09,9E+09,9E+09,9E+09,9E+09]];
    CONST robtarget Target_70NomLab_I:=[[-39.178192,-12.698133,-20],[0.707106781,0,0,0.707106781],[0,0,0,0],[9E+09,9E+09,9E+09,9E+09,9E+09,9E+09]];
    CONST robtarget Target_150NomLab_R:=[[-53.243442,-12.562931,-20],[0.707106781,0,0,0.707106781],[0,0,0,0],[9E+09,9E+09,9E+09,9E+09,9E+09,9E+09]];
    CONST robtarget Target_80NomLab_Rint:=[[-87.50619,-27.43225,-20],[0.707106781,0,0,0.707106781],[0,0,0,0],[9E+09,9E+09,9E+09,9E+09,9E+09,9E+09]];
    CONST robtarget Target_Nom_L_100:=[[3.79755,47.324448,-20],[0.707106781,0,0,0.707106781],[0,0,0,0],[9E+09,9E+09,9E+09,9E+09,9E+09,9E+09]];
    CONST robtarget Target_Nom_L_20:=[[3.79755,47.324448,0],[0.707106781,0,0,0.707106781],[0,0,0,0],[9E+09,9E+09,9E+09,9E+09,9E+09,9E+09]];
    CONST robtarget Target_Nom_L_30:=[[2.597069625,3.348416,0],[0.707106781,0,0,0.707106781],[0,0,0,0],[9E+09,9E+09,9E+09,9E+09,9E+09,9E+09]];
    CONST robtarget Target_Nom_L_40:=[[-1.998180875,0.1710675,0],[0.707106781,0,0,0.707106781],[0,0,0,0],[9E+09,9E+09,9E+09,9E+09,9E+09,9E+09]];
    CONST robtarget Target_Nom_L_50:=[[-9.708635,-0.116667,0],[0.707106781,0,0,0.707106781],[0,0,0,0],[9E+09,9E+09,9E+09,9E+09,9E+09,9E+09]];
    CONST robtarget Target_Nom_L_60:=[[-9.708635,5.12076,0],[0.707106781,0,0,0.707106781],[0,0,0,0],[9E+09,9E+09,9E+09,9E+09,9E+09,9E+09]];
    CONST robtarget Target_Nom_L_70:=[[-1.286154,6.56909,0],[0.707106781,0,0,0.707106781],[0,0,0,0],[9E+09,9E+09,9E+09,9E+09,9E+09,9E+09]];
    CONST robtarget Target_Nom_L_80:=[[-1.286154,47.476319,0],[0.707106781,0,0,0.707106781],[0,0,0,0],[9E+09,9E+09,9E+09,9E+09,9E+09,9E+09]];
    CONST robtarget Target_Nom_L_90:=[[3.79755,47.324448,0],[0.707106781,0,0,0.707106781],[0,0,0,0],[9E+09,9E+09,9E+09,9E+09,9E+09,9E+09]];
    CONST robtarget Target_Nom_L_10:=[[3.79755,47.324448,-20],[0.707106781,0,0,0.707106781],[0,0,0,0],[9E+09,9E+09,9E+09,9E+09,9E+09,9E+09]];
    CONST robtarget Target_Nom_A_10:=[[-44.486792,29.956669,-20],[0.707106781,0,0,0.707106781],[0,0,0,0],[9E+09,9E+09,9E+09,9E+09,9E+09,9E+09]];
    CONST robtarget Target_Nom_A_20:=[[-44.486792,29.956669,0],[0.707106781,0,0,0.707106781],[0,0,0,0],[9E+09,9E+09,9E+09,9E+09,9E+09,9E+09]];
    CONST robtarget Target_Nom_A_30:=[[-45.446965,20.377958,0],[0.707106781,0,0,0.707106781],[0,-1,0,0],[9E+09,9E+09,9E+09,9E+09,9E+09,9E+09]];
    CONST robtarget Target_Nom_A_40:=[[-14.033515,20.377958,0],[0.707106781,0,0,0.707106781],[0,-1,0,0],[9E+09,9E+09,9E+09,9E+09,9E+09,9E+09]];
    CONST robtarget Target_Nom_A_50:=[[-14.912725,3.965854,0],[0.707106781,0,0,0.707106781],[0,-1,0,0],[9E+09,9E+09,9E+09,9E+09,9E+09,9E+09]];
    CONST robtarget Target_Nom_A_60:=[[-19.425723,0.264069,0],[0.707106781,0,0,0.707106781],[0,-1,0,0],[9E+09,9E+09,9E+09,9E+09,9E+09,9E+09]];
    CONST robtarget Target_Nom_A_70:=[[-50.454998,-0.116667,0],[0.707106781,0,0,0.707106781],[0,-1,0,0],[9E+09,9E+09,9E+09,9E+09,9E+09,9E+09]];
    CONST robtarget Target_Nom_A_80:=[[-49.995417,30.69565,0],[0.707106781,0,0,0.707106781],[0,-1,0,0],[9E+09,9E+09,9E+09,9E+09,9E+09,9E+09]];
    CONST robtarget Target_Nom_A_90:=[[-45.087396,35.436719,0],[0.707106781,0,0,0.707106781],[0,-1,0,0],[9E+09,9E+09,9E+09,9E+09,9E+09,9E+09]];
    CONST robtarget Target_Nom_A_100:=[[-14.033515,35.635156,0],[0.707106781,0,0,0.707106781],[0,-1,0,0],[9E+09,9E+09,9E+09,9E+09,9E+09,9E+09]];
    CONST robtarget Target_Nom_A_110:=[[-14.033515,30.625271,0],[0.707106781,0,0,0.707106781],[0,-1,0,0],[9E+09,9E+09,9E+09,9E+09,9E+09,9E+09]];
    CONST robtarget Target_Nom_A_120:=[[-44.486792,29.956669,0],[0.707106781,0,0,0.707106781],[0,-1,0,0],[9E+09,9E+09,9E+09,9E+09,9E+09,9E+09]];
    CONST robtarget Target_Nom_A_130:=[[-44.486792,29.956669,-20],[0.707106781,0,0,0.707106781],[0,-1,0,0],[9E+09,9E+09,9E+09,9E+09,9E+09,9E+09]];
    CONST robtarget Target_Nom_Aint_10:=[[-45.191377,15.060362,-20],[0.707106781,0,0,0.707106781],[0,0,0,0],[9E+09,9E+09,9E+09,9E+09,9E+09,9E+09]];
    CONST robtarget Target_Nom_Aint_20:=[[-45.191377,15.060362,0],[0.707106781,0,0,0.707106781],[0,0,0,0],[9E+09,9E+09,9E+09,9E+09,9E+09,9E+09]];
    CONST robtarget Target_Nom_Aint_30:=[[-45.333194,5.234796,0],[0.707106781,0,0,0.707106781],[0,0,0,0],[9E+09,9E+09,9E+09,9E+09,9E+09,9E+09]];
    CONST robtarget Target_Nom_Aint_40:=[[-20.275035,5.361796,0],[0.707106781,0,0,0.707106781],[0,0,0,0],[9E+09,9E+09,9E+09,9E+09,9E+09,9E+09]];
    CONST robtarget Target_Nom_Aint_50:=[[-19.041548,15.342144,0],[0.707106781,0,0,0.707106781],[0,0,0,0],[9E+09,9E+09,9E+09,9E+09,9E+09,9E+09]];
    CONST robtarget Target_Nom_Aint_60:=[[-45.191377,15.060362,0],[0.707106781,0,0,0.707106781],[0,0,0,0],[9E+09,9E+09,9E+09,9E+09,9E+09,9E+09]];
    CONST robtarget Target_Nom_Aint_70:=[[-45.191377,15.060362,-20],[0.707106781,0,0,0.707106781],[0,0,0,0],[9E+09,9E+09,9E+09,9E+09,9E+09,9E+09]];
    CONST robtarget Target_Nom_B_10:=[[-70.800398,-0.116667,-20],[0.707106781,0,0,0.707106781],[0,-1,0,0],[9E+09,9E+09,9E+09,9E+09,9E+09,9E+09]];
    CONST robtarget Target_Nom_B_20:=[[-70.800398,-0.116667,0],[0.707106781,0,0,0.707106781],[0,0,0,0],[9E+09,9E+09,9E+09,9E+09,9E+09,9E+09]];
    CONST robtarget Target_Nom_B_30:=[[-88.365821,0.91071,0],[0.707106781,0,0,0.707106781],[0,0,0,0],[9E+09,9E+09,9E+09,9E+09,9E+09,9E+09]];
    CONST robtarget Target_Nom_B_40:=[[-92.0476305,7.729816625,0],[0.707106781,0,0,0.707106781],[0,0,0,0],[9E+09,9E+09,9E+09,9E+09,9E+09,9E+09]];
    CONST robtarget Target_Nom_B_50:=[[-90.973554,32.296115,0],[0.707106781,0,0,0.707106781],[0,0,0,0],[9E+09,9E+09,9E+09,9E+09,9E+09,9E+09]];
    CONST robtarget Target_Nom_B_60:=[[-87.050048,35.424019,0],[0.707106781,0,0,0.707106781],[0,0,0,0],[9E+09,9E+09,9E+09,9E+09,9E+09,9E+09]];
    CONST robtarget Target_Nom_B_70:=[[-60.760221375,36.8803515,0],[0.707106781,0,0,0.707106781],[0,0,0,0],[9E+09,9E+09,9E+09,9E+09,9E+09,9E+09]];
    CONST robtarget Target_Nom_B_80:=[[-60.698342,47.476319,0],[0.707106781,0,0,0.707106781],[0,0,0,0],[9E+09,9E+09,9E+09,9E+09,9E+09,9E+09]];
    CONST robtarget Target_Nom_B_90:=[[-55.690573,47.476319,0],[0.707106781,0,0,0.707106781],[0,0,0,0],[9E+09,9E+09,9E+09,9E+09,9E+09,9E+09]];
    CONST robtarget Target_Nom_B_100:=[[-55.690573,-0.116667,0],[0.707106781,0,0,0.707106781],[0,0,0,0],[9E+09,9E+09,9E+09,9E+09,9E+09,9E+09]];
    CONST robtarget Target_Nom_B_110:=[[-70.800398,-0.116667,0],[0.707106781,0,0,0.707106781],[0,0,0,0],[9E+09,9E+09,9E+09,9E+09,9E+09,9E+09]];
    CONST robtarget Target_Nom_B_120:=[[-70.800398,-0.116667,-20],[0.707106781,0,0,0.707106781],[0,0,0,0],[9E+09,9E+09,9E+09,9E+09,9E+09,9E+09]];
    CONST robtarget Target_Nom_Bint_10:=[[-86.202058,29.967252,-20],[0.707106781,0,0,0.707106781],[0,0,0,0],[9E+09,9E+09,9E+09,9E+09,9E+09,9E+09]];
    CONST robtarget Target_Nom_Bint_20:=[[-86.202058,29.967252,0],[0.707106781,0,0,0.707106781],[0,0,0,0],[9E+09,9E+09,9E+09,9E+09,9E+09,9E+09]];
    CONST robtarget Target_Nom_Bint_30:=[[-86.321385,5.818996,0],[0.707106781,0,0,0.707106781],[0,0,0,0],[9E+09,9E+09,9E+09,9E+09,9E+09,9E+09]];
    CONST robtarget Target_Nom_Bint_40:=[[-61.534425,5.843338,0],[0.707106781,0,0,0.707106781],[0,0,0,0],[9E+09,9E+09,9E+09,9E+09,9E+09,9E+09]];
    CONST robtarget Target_Nom_Bint_50:=[[-61.592898,29.928094,0],[0.707106781,0,0,0.707106781],[0,0,0,0],[9E+09,9E+09,9E+09,9E+09,9E+09,9E+09]];
    CONST robtarget Target_Nom_Bint_60:=[[-86.202058,29.967252,0],[0.707106781,0,0,0.707106781],[0,0,0,0],[9E+09,9E+09,9E+09,9E+09,9E+09,9E+09]];
    CONST robtarget Target_Nom_Bint_70:=[[-86.202058,29.967252,-20],[0.707106781,0,0,0.707106781],[0,0,0,0],[9E+09,9E+09,9E+09,9E+09,9E+09,9E+09]];
    CONST robtarget Target_Nom_S_250:=[[3.133975,-12.610292,-20],[0.707106781,0,0,0.707106781],[0,0,0,0],[9E+09,9E+09,9E+09,9E+09,9E+09,9E+09]];
    CONST robtarget Target_Nom_S_240:=[[3.133975,-12.610292,0],[0.707106781,0,0,0.707106781],[0,0,0,0],[9E+09,9E+09,9E+09,9E+09,9E+09,9E+09]];
    CONST robtarget Target_Nom_S_30:=[[10.437004,-18.903406,0],[0.707106781,0,0,0.707106781],[0,0,0,0],[9E+09,9E+09,9E+09,9E+09,9E+09,9E+09]];
    CONST robtarget Target_Nom_S_40:=[[9.772106,-34.450058,0],[0.707106781,0,0,0.707106781],[0,0,0,0],[9E+09,9E+09,9E+09,9E+09,9E+09,9E+09]];
    CONST robtarget Target_Nom_S_50:=[[4.860117,-38.959088,0],[0.707106781,0,0,0.707106781],[0,0,0,0],[9E+09,9E+09,9E+09,9E+09,9E+09,9E+09]];
    CONST robtarget Target_Nom_S_60:=[[-23.935546,-39.625838,0],[0.707106781,0,0,0.707106781],[0,0,0,0],[9E+09,9E+09,9E+09,9E+09,9E+09,9E+09]];
    CONST robtarget Target_Nom_S_70:=[[-23.935546,-47.140533,0],[0.707106781,0,0,0.707106781],[0,0,0,0],[9E+09,9E+09,9E+09,9E+09,9E+09,9E+09]];
    CONST robtarget Target_Nom_S_80:=[[0.973917,-47.368075,0],[0.707106781,0,0,0.707106781],[0,0,0,0],[9E+09,9E+09,9E+09,9E+09,9E+09,9E+09]];
    CONST robtarget Target_Nom_S_90:=[[1.104092,-43.724763,0],[0.707106781,0,0,0.707106781],[0,0,0,0],[9E+09,9E+09,9E+09,9E+09,9E+09,9E+09]];
    CONST robtarget Target_Nom_S_100:=[[10.550775,-43.601467,0],[0.707106781,0,0,0.707106781],[0,0,0,0],[9E+09,9E+09,9E+09,9E+09,9E+09,9E+09]];
    CONST robtarget Target_Nom_S_110:=[[8.714037,-53.402692,0],[0.707106781,0,0,0.707106781],[0,0,0,0],[9E+09,9E+09,9E+09,9E+09,9E+09,9E+09]];
    CONST robtarget Target_Nom_S_120:=[[2.923631,-56.786713,0],[0.707106781,0,0,0.707106781],[0,0,0,0],[9E+09,9E+09,9E+09,9E+09,9E+09,9E+09]];
    CONST robtarget Target_Nom_S_130:=[[-26.667104,-56.674,0],[0.707106781,0,0,0.707106781],[0,0,0,0],[9E+09,9E+09,9E+09,9E+09,9E+09,9E+09]];
    CONST robtarget Target_Nom_S_140:=[[-32.793233875,-51.677079125,0],[0.707106781,0,0,0.707106781],[0,0,0,0],[9E+09,9E+09,9E+09,9E+09,9E+09,9E+09]];
    CONST robtarget Target_Nom_S_150:=[[-32.840263125,-35.198696625,0],[0.707106781,0,0,0.707106781],[0,0,0,0],[9E+09,9E+09,9E+09,9E+09,9E+09,9E+09]];
    CONST robtarget Target_Nom_S_160:=[[-26.023637,-29.974631,0],[0.707106781,0,0,0.707106781],[0,0,0,0],[9E+09,9E+09,9E+09,9E+09,9E+09,9E+09]];
    CONST robtarget Target_Nom_S_170:=[[0.990321,-29.720102,0],[0.707106781,0,0,0.707106781],[0,0,0,0],[9E+09,9E+09,9E+09,9E+09,9E+09,9E+09]];
    CONST robtarget Target_Nom_S_180:=[[0.990585,-22.091371,0],[0.707106781,0,0,0.707106781],[0,0,0,0],[9E+09,9E+09,9E+09,9E+09,9E+09,9E+09]];
    CONST robtarget Target_Nom_S_190:=[[-23.979532875,-22.814046875,0],[0.707106781,0,0,0.707106781],[0,0,0,0],[9E+09,9E+09,9E+09,9E+09,9E+09,9E+09]];
    CONST robtarget Target_Nom_S_200:=[[-24.049317,-25.848719,0],[0.707106781,0,0,0.707106781],[0,0,0,0],[9E+09,9E+09,9E+09,9E+09,9E+09,9E+09]];
    CONST robtarget Target_Nom_S_210:=[[-33.837577,-25.848719,0],[0.707106781,0,0,0.707106781],[0,0,0,0],[9E+09,9E+09,9E+09,9E+09,9E+09,9E+09]];
    CONST robtarget Target_Nom_S_220:=[[-31.20606425,-15.42115925,0],[0.707106781,0,0,0.707106781],[0,0,0,0],[9E+09,9E+09,9E+09,9E+09,9E+09,9E+09]];
    CONST robtarget Target_Nom_S_230:=[[-25.843456,-12.413442,0],[0.707106781,0,0,0.707106781],[0,0,0,0],[9E+09,9E+09,9E+09,9E+09,9E+09,9E+09]];
    CONST robtarget Target_Nom_S_20:=[[3.133975,-12.610292,0],[0.707106781,0,0,0.707106781],[0,0,0,0],[9E+09,9E+09,9E+09,9E+09,9E+09,9E+09]];
    CONST robtarget Target_Nom_S_10:=[[3.133975,-12.610292,-20],[0.707106781,0,0,0.707106781],[0,0,0,0],[9E+09,9E+09,9E+09,9E+09,9E+09,9E+09]];
    CONST robtarget Target_Nom_I_10:=[[-39.178192,-12.698133,-20],[0.707106781,0,0,0.707106781],[0,0,0,0],[9E+09,9E+09,9E+09,9E+09,9E+09,9E+09]];
    CONST robtarget Target_Nom_I_20:=[[-39.178192,-12.698133,0],[0.707106781,0,0,0.707106781],[0,0,0,0],[9E+09,9E+09,9E+09,9E+09,9E+09,9E+09]];
    CONST robtarget Target_Nom_I_30:=[[-39.186923,-56.932233,0],[0.707106781,0,0,0.707106781],[0,0,0,0],[9E+09,9E+09,9E+09,9E+09,9E+09,9E+09]];
    CONST robtarget Target_Nom_I_40:=[[-48.633871,-57.055529,0],[0.707106781,0,0,0.707106781],[0,0,0,0],[9E+09,9E+09,9E+09,9E+09,9E+09,9E+09]];
    CONST robtarget Target_Nom_I_50:=[[-48.633871,-12.413442,0],[0.707106781,0,0,0.707106781],[0,0,0,0],[9E+09,9E+09,9E+09,9E+09,9E+09,9E+09]];
    CONST robtarget Target_Nom_I_60:=[[-39.178192,-12.698133,0],[0.707106781,0,0,0.707106781],[0,0,0,0],[9E+09,9E+09,9E+09,9E+09,9E+09,9E+09]];
    CONST robtarget Target_Nom_I_70:=[[-39.178192,-12.698133,-20],[0.707106781,0,0,0.707106781],[0,0,0,0],[9E+09,9E+09,9E+09,9E+09,9E+09,9E+09]];
    CONST robtarget Target_Nom_R_150:=[[-53.243442,-12.562931,-20],[0.707106781,0,0,0.707106781],[0,0,0,0],[9E+09,9E+09,9E+09,9E+09,9E+09,9E+09]];
    CONST robtarget Target_Nom_R_140:=[[-53.243442,-12.562931,0],[0.707106781,0,0,0.707106781],[0,0,0,0],[9E+09,9E+09,9E+09,9E+09,9E+09,9E+09]];
    CONST robtarget Target_Nom_R_30:=[[-52.95875,-57.055529,0],[0.707106781,0,0,0.707106781],[0,0,0,0],[9E+09,9E+09,9E+09,9E+09,9E+09,9E+09]];
    CONST robtarget Target_Nom_R_40:=[[-62.405698,-56.932233,0],[0.707106781,0,0,0.707106781],[0,0,0,0],[9E+09,9E+09,9E+09,9E+09,9E+09,9E+09]];
    CONST robtarget Target_Nom_R_50:=[[-62.525819,-42.543663,0],[0.707106781,0,0,0.707106781],[0,0,0,0],[9E+09,9E+09,9E+09,9E+09,9E+09,9E+09]];
    CONST robtarget Target_Nom_R_60:=[[-76.007133,-43.470763,0],[0.707106781,0,0,0.707106781],[0,0,0,0],[9E+09,9E+09,9E+09,9E+09,9E+09,9E+09]];
    CONST robtarget Target_Nom_R_70:=[[-87.563869,-57.055265,0],[0.707106781,0,0,0.707106781],[0,0,0,0],[9E+09,9E+09,9E+09,9E+09,9E+09,9E+09]];
    CONST robtarget Target_Nom_R_80:=[[-97.233596,-56.932233,0],[0.707106781,0,0,0.707106781],[0,0,0,0],[9E+09,9E+09,9E+09,9E+09,9E+09,9E+09]];
    CONST robtarget Target_Nom_R_90:=[[-95.014006,-50.87645,0],[0.707106781,0,0,0.707106781],[0,0,0,0],[9E+09,9E+09,9E+09,9E+09,9E+09,9E+09]];
    CONST robtarget Target_Nom_R_100:=[[-88.582646625,-42.2683965,0],[0.707106781,0,0,0.707106781],[0,0,0,0],[9E+09,9E+09,9E+09,9E+09,9E+09,9E+09]];
    CONST robtarget Target_Nom_R_110:=[[-96.168912,-37.385346,0],[0.707106781,0,0,0.707106781],[0,0,0,0],[9E+09,9E+09,9E+09,9E+09,9E+09,9E+09]];
    CONST robtarget Target_Nom_R_120:=[[-96.036725312,-17.219842617,0],[0.707106781,0,0,0.707106781],[0,0,0,0],[9E+09,9E+09,9E+09,9E+09,9E+09,9E+09]];
    CONST robtarget Target_Nom_R_130:=[[-91.922615,-13.372292,0],[0.707106781,0,0,0.707106781],[0,0,0,0],[9E+09,9E+09,9E+09,9E+09,9E+09,9E+09]];
    CONST robtarget Target_Nom_R_20:=[[-53.243442,-12.562931,0],[0.707106781,0,0,0.707106781],[0,0,0,0],[9E+09,9E+09,9E+09,9E+09,9E+09,9E+09]];
    CONST robtarget Target_Nom_R_10:=[[-53.243442,-12.562931,-20],[0.707106781,0,0,0.707106781],[0,0,0,0],[9E+09,9E+09,9E+09,9E+09,9E+09,9E+09]];
    CONST robtarget Target_Nom_Rint_10:=[[-87.50619,-27.43225,-20],[0.707106781,0,0,0.707106781],[0,0,0,0],[9E+09,9E+09,9E+09,9E+09,9E+09,9E+09]];
    CONST robtarget Target_Nom_Rint_20:=[[-87.50619,-27.43225,0],[0.707106781,0,0,0.707106781],[0,0,0,0],[9E+09,9E+09,9E+09,9E+09,9E+09,9E+09]];
    CONST robtarget Target_Nom_Rint_30:=[[-87.567573,-32.68026,0],[0.707106781,0,0,0.707106781],[0,0,0,0],[9E+09,9E+09,9E+09,9E+09,9E+09,9E+09]];
